  def set_closed_mm(closed_mm, gripper_socket):
      gripper_closed_mm[to_num(gripper_socket) - 1] = closed_mm
  end

  def set_open_mm(open_mm, gripper_socket):
      gripper_open_mm[to_num(gripper_socket) - 1] = open_mm
  end

  def gripper_to_mm(value_gripper, gripper_socket):
      closed_norm = get_closed_norm(gripper_socket)
      open_norm = get_open_norm(gripper_socket)
      closed_mm = get_closed_mm(gripper_socket)
      open_mm = get_open_mm(gripper_socket)

      value_norm = (value_gripper / 255) * 100

      slope = (closed_mm - open_mm) / (closed_norm - open_norm)
      value_mm = slope * (value_norm - closed_norm) + closed_mm

      if (value_mm > open_mm):
          value_mm_limited = open_mm
      elif (value_mm < closed_mm):
          value_mm_limited = closed_mm
      else:
          value_mm_limited = value_mm
      end

      return value_mm_limited
  end

  def mm_to_gripper(value_mm, gripper_socket):
      closed_norm = get_closed_norm(gripper_socket)
      open_norm = get_open_norm(gripper_socket)
      closed_mm = get_closed_mm(gripper_socket)
      open_mm = get_open_mm(gripper_socket)

      slope = (closed_norm - open_norm) / (closed_mm - open_mm)
      value_norm = (value_mm - closed_mm) * slope + closed_norm

      value_gripper = value_norm * 255 / 100

      if (value_gripper > 255):
          value_gripper_limited = 255
      elif (value_gripper < 0):
          value_gripper_limited = 0
      else:
          value_gripper_limited = round_value(value_gripper)
      end

      return value_gripper_limited
  end

  def round_value(value):
      value_mod = value % 1

      if(value_mod < 0.5):
          return floor(value)
      else:
          return ceil(value)
      end
  end

  def round_value_2_dec(value):
      value_x_100 = value * 100
      value_x_100_rounded = round_value(value_x_100)
      return value_x_100_rounded / 100
  end

  def clear_socket_buffer(gripper_socket="1", read_timeout = 0.1):
      rq_comm_clear_socket_buffer_enabled[rq_socket_to_index(gripper_socket)] = True
  end

  def rq_gripper_id_to_ascii(gripper_id):
      if(gripper_id == "1"):
          return 57
      elif(gripper_id == "2"):
          return 50
      elif(gripper_id == "3"):
          return 51
      elif(gripper_id == "4"):
          return 52
      end
  end

      def scale(value, rawRange, scaledRange):
          def computeSlope(inputRange, outputRange):
              outputRangeDelta = outputRange[1] - outputRange[0]
              inputRangeDelta = inputRange[1] - inputRange[0]

              if (inputRangeDelta == 0):
                  return 0
              else:
                  return outputRangeDelta / inputRangeDelta
              end
          end

          def computeIntercept(slope, inputRange, outputRange):
              return outputRange[0] - (slope * inputRange[0])
          end

          def clipScaledValue(outputScaledValue, outputRange):
              if (outputRange[0] < outputRange[1]):
                  return clipWhenLowerLimitIsLessThanHigher(outputScaledValue, outputRange)
              else:
                  return clipWhenLowerLimitIsGreaterThanHigherLimit(outputScaledValue, outputRange)
              end
          end

          def clipWhenLowerLimitIsGreaterThanHigherLimit(outputScaledValue, outputRange):
              if (outputScaledValue < outputRange[1]):
                  return outputRange[1]
              elif (outputScaledValue > outputRange[0]):
                  return outputRange[0]
              else:
                  return outputScaledValue
              end
          end

          def clipWhenLowerLimitIsLessThanHigher(outputScaledValue, outputRange):
              if (outputScaledValue < outputRange[0]):
                  return outputRange[0]
              elif (outputScaledValue > outputRange[1]):
                  return outputRange[1]
              else:
                  return outputScaledValue
              end
          end

          slope = computeSlope(rawRange, scaledRange)
          intercept = computeIntercept(slope, rawRange, scaledRange)
          scaledValue = slope * value + intercept
          return clipScaledValue(scaledValue, scaledRange)
      end

      def limit(value, range):
          return scale(value, range, range)
      end


  rq_init_comm_if_connected(9, "1")
  rq_init_comm_if_connected(2, "2")
  rq_init_comm_if_connected(3, "3")
  rq_init_comm_if_connected(4, "4")
  rq_print_connected_grippers()
  rq_gripper_communication_thread = run rq_gripper_communication()
  set_closed_norm(97.6470588235294, "1")
  set_open_norm(1.1764705882352942, "1")
  set_closed_mm(0.0, "1")
  set_open_mm(53.0, "1")
  set_closed_norm(100.0, "2")
  set_open_norm(0.0, "2")
  set_closed_mm(0.0, "2")
  set_open_mm(50.0, "2")
  set_closed_norm(100.0, "3")
  set_open_norm(0.0, "3")
  set_closed_mm(0.0, "3")
  set_open_mm(50.0, "3")
  set_closed_norm(100.0, "4")
  set_open_norm(0.0, "4")
  set_closed_mm(0.0, "4")
  set_open_mm(50.0, "4")
  rq_current_limit_enabled = False
  while(not rq_gripper_communication_thread_started):
      sleep(0.008)
  end
  # end: URCap Installation Node
  global AMR_Position=struct(position_identifier=0, x1=0, x2=0, y1=0, y2=0, theta1=0, theta2=0)
  global CAM_Pose=p[0,0,0,0,0,0]
  global CAM_Relation=""
  global CMD_Abort=  False
  global CMD_Clear=  False
  global CMD_Reset=  False
  global CMD_Start=  False
  global CMD_Suspend=  False
  global CMD_Unhold=  False
  global CMD_Unsuspend=  False
  global CNT_Rack_Output=0
  global FNC_Freedrive=  False
  global PRC_TubCounter=0
  global STP=0
  global easyPickCount_4=0
  global easyPickCount_7=0
  global easyPickNoObj_4=0
  global easyPickNoObj_7=0
  global easyPickParts_4=0
  global easyPickParts_7=0
  global TMR_Barcode=0
  global Container_mid_1_p=p[-.379239199143, -.127191311915, .299999999998, .000000000046, -.000000000021, -1.247199999994]
  global Container_mid_1_q=[-2.477408934449926, -1.2969853503591224, -1.875639182904262, -1.539621866126728, 1.5731943360401213, -2.8009955944022717]
  global trigger_otw_p=p[-.364831738276, -.163967193938, .343299997821, .000000000046, -.000000000020, -1.148401333327]
  global trigger_otw_q=[-2.378283213085033, -1.2994862387706814, -1.7634300687554951, -1.6493302004167063, 1.573123683454141, -2.8011223671816943]
  global Waypoint_54_p=p[.008800512419, -.547926542621, .402696567415, -.589884378425, -.007228654778, -.061268144704]
  global Waypoint_54_q=[-1.2044575850116175, -1.3416667741588135, -1.8272563219070435, -0.9884541195682068, 1.3621035814285278, -2.7712565104113978]
  global Waypoint_77_p=p[-.178371829612, -.433927395311, .368082383916, -.086593488055, .704679941724, -.007869906074]
  global Waypoint_77_q=[-1.265390698109762, -1.3355963987163086, -1.7944865226745605, -1.7402602634825648, 0.8780410885810852, -2.7713127771960657]
  global Waypoint_83_p=p[.008800512419, -.547926542621, .402696567415, -.589884378425, -.007228654778, -.061268144704]
  global Waypoint_83_q=[-1.2044575850116175, -1.3416667741588135, -1.8272563219070435, -0.9884541195682068, 1.3621035814285278, -2.7712565104113978]
  global Waypoint_84_p=p[-.178371829612, -.433927395311, .368082383916, -.086593488055, .704679941724, -.007869906074]
  global Waypoint_84_q=[-1.265390698109762, -1.3355963987163086, -1.7944865226745605, -1.7402602634825648, 0.8780410885810852, -2.7713127771960657]
  global Vial_above_1_p=p[.017105793010, -.652093028359, .184920586844, .000000000272, .000000000270, 1.564063451276]
  global Vial_above_1_q=[-1.3375440709712851, -1.9618096977868804, -1.4665759083780685, -1.2837941559171444, 1.5732503672317195, -4.47276330421513]
  global Vial_pick_poi_1_p=p[.017105792852, -.648922724010, .093307568731, .000000000271, .000000000270, 1.564063451276]
  global Vial_pick_poi_1_q=[-1.3366329456391917, -2.0375277831965413, -1.6071432798879028, -1.0675084332049813, 1.57309887265915, -4.471135348858068]
  global Waypoint_86_p=p[.019227646885, -.648669633640, .184920586950, .000000000000, .000000000000, .024063451426]
  global Waypoint_86_q=[-1.3331129109407733, -1.9540750545686123, -1.4775914902901128, -1.280581784992414, 1.5733500744865856, -2.928303704452631]
  global Waypoint_87_p=p[-.032361834699, -.348336136197, .391475576335, -.000008499254, .000014589902, -.004651426820]
  global Waypoint_87_q=[-1.2709335019096129, -1.1914598663441005, -1.708995335060501, -1.8117888533498316, 1.5729683532263925, -2.8379347397710237]
  global Vial_3FG_plac_1_p=p[-.031858676359, -.349402499566, .145301120695, .000000000000, .000000000000, .000000000000]
  global Vial_3FG_plac_1_q=[-1.2723975525801707, -1.252376585823825, -2.3128114007049496, -1.1470592278900167, 1.5730548099411423, -2.8414815174610535]
  global Waypoint_88_p=p[-.032361834699, -.348336136197, .391475576335, -.000008499254, .000014589902, -.004651426820]
  global Waypoint_88_q=[-1.2709335019096129, -1.1914598663441005, -1.708995335060501, -1.8117888533498316, 1.5729683532263925, -2.8379347397710237]
  global cap_dump_1_p=p[-.139168676487, -.420163541420, .146096395183, .000000000000, .000000000000, .000000000000]
  global cap_dump_1_q=[-1.584588644510994, -1.5093464179777323, -2.1118449369620347, -1.091059703602438, 1.5728943834877336, -3.154014906686923]
  global Waypoint_89_p=p[-.032361834699, -.348336136197, .391475576335, -.000008499254, .000014589902, -.004651426820]
  global Waypoint_89_q=[-1.2709335019096129, -1.1914598663441005, -1.708995335060501, -1.8117888533498316, 1.5729683532263925, -2.8379347397710237]
  global Vial_3FG_plac_2_p=p[-.031858676359, -.349402499566, .145301120695, .000000000000, .000000000000, .000000000000]
  global Vial_3FG_plac_2_q=[-1.2723975525801707, -1.252376585823825, -2.3128114007049496, -1.1470592278900167, 1.5730548099411423, -2.8414815174610535]
  global Waypoint_90_p=p[-.032361834699, -.348336136197, .391475576335, -.000008499254, .000014589902, -.004651426820]
  global Waypoint_90_q=[-1.2709335019096129, -1.1914598663441005, -1.708995335060501, -1.8117888533498316, 1.5729683532263925, -2.8379347397710237]
  global cap_dump_2_p=p[-.139168676487, -.420163541420, .146096395183, .000000000000, .000000000000, .000000000000]
  global cap_dump_2_q=[-1.584588644510994, -1.5093464179777323, -2.1118449369620347, -1.091059703602438, 1.5728943834877336, -3.154014906686923]
  global Waypoint_91_p=p[-.032361834699, -.348336136197, .391475576335, -.000008499254, .000014589902, -.004651426820]
  global Waypoint_91_q=[-1.2709335019096129, -1.1914598663441005, -1.708995335060501, -1.8117888533498316, 1.5729683532263925, -2.8379347397710237]
  global Vial_liq_abov_1_p=p[-.025303660977, -.338758622354, .426628485936, -1.315858642253, .800043520260, -.928295855026]
  global Vial_liq_abov_1_q=[-0.3789628187762659, -1.5149522957256814, -2.263045310974121, 0.7870649534412841, -0.750984017048971, -3.2237566153155726]
  global Vial_liq_pick_3_p=p[-.002660428945, -.335984893034, .159389832934, -1.150456778400, .673175527684, -1.010612657503]
  global Vial_liq_pick_3_q=[-0.3660772482501429, -1.4503649038127442, -2.4056053161621094, -1.994692941705221, 0.8039668202400208, -0.2508929411517542]
  global Vial_liq_pick_4_p=p[-.041402486291, -.356791603314, .125395323246, -1.143483969075, .651070210027, -.878721885453]
  global Vial_liq_pick_4_q=[-0.4426233705502476, -1.437252121513727, -2.551930962114307, -1.776528229806984, 0.6562026234073748, -0.43018811960029524]
  global Vial_liq_abov_2_p=p[-.025303660977, -.338758622354, .426628485936, -1.315858642253, .800043520260, -.928295855026]
  global Vial_liq_abov_2_q=[-0.3789628187762659, -1.5149522957256814, -2.263045310974121, 0.7870649534412841, -0.750984017048971, -3.2237566153155726]
  global Liquid_midway_1_p=p[.057575295009, -.583081747994, .306414980749, -1.351675548728, .120935756539, -.096908606303]
  global Liquid_midway_1_q=[-0.895174805318014, -1.7035466633238734, -2.380953073501587, 0.631549521083496, 0.7706599235534668, -2.9455552736865442]
  global shake_3_p=p[.057574880217, -.583085370269, .306422893466, -1.360996190983, -.155555042453, -.438136255921]
  global shake_3_q=[-0.8951800505267542, -1.7035466633238734, -2.380937099456787, 0.6315542894550782, 0.7706599235534669, -2.5394540616517496]
  global shake_4_p=p[.057581636113, -.583090570002, .306439684073, -1.308767904323, .368530312677, .214926493520]
  global shake_4_q=[-0.8951714674579065, -1.7035395107665003, -2.380906343460083, 0.6315504747578125, 0.7706480026245118, -3.3161255787892268]
  global drop_above_3_p=p[.268235025993, -.467784390499, .226219872376, -1.027832627524, -.430841408251, 1.004603115937]
  global drop_above_3_q=[-0.935645882283346, -1.6663371525206507, -2.4252893924713135, 0.41966931402172847, 1.8470635414123535, -3.4600217978106897]
  global drop_above_4_p=p[.219042229014, -.470775657081, .133754190740, -.313004595901, -.344395319364, 1.500564994056]
  global drop_above_4_q=[-1.0601594887284795, -1.70046459045642, -2.0799996233759863, -0.7243227230676759, 1.9429634314685202, -4.115129153870795]
  global liq_tran_3_p=p[.213067510942, -.469567035397, .100231043184, .251862243732, .217902579404, 1.592812335393]
  global liq_tran_3_q=[-0.7789645168037476, -1.822364827406652, -1.8643518410805573, -1.252158963840138, 1.3768134449520435, -3.9328333233290254]
  global drop_above_5_p=p[.219042229014, -.470775657081, .133754190740, -.313004595901, -.344395319364, 1.500564994056]
  global drop_above_5_q=[-1.0601594887284795, -1.70046459045642, -2.0799996233759863, -0.7243227230676759, 1.9429634314685202, -4.115129153870795]
  global Waypoint_92_p=p[.187119460405, -.493959476151, .133754190608, -.313004596540, -.344395317757, 1.500564993991]
  global Waypoint_92_q=[-1.1418328121400876, -1.7310553375189475, -2.033634768766424, -0.772026910513711, 1.958578934631971, -4.201588449364511]
  global liq_tran_4_p=p[.195957706507, -.493022614126, .100231042689, .160718757180, .109807038912, 1.525321508623]
  global liq_tran_4_q=[-0.881740380645474, -1.8244526267589851, -1.865100964490387, -1.1608866323693583, 1.4631433601076713, -3.973915130363038]
  global drop_above_6_p=p[.219042229014, -.470775657081, .133754190740, -.313004595901, -.344395319364, 1.500564994056]
  global drop_above_6_q=[-1.0601594887284795, -1.70046459045642, -2.0799996233759863, -0.7243227230676759, 1.9429634314685202, -4.115129153870795]
  global drop_above_7_p=p[.268235025993, -.467784390499, .226219872376, -1.027832627524, -.430841408251, 1.004603115937]
  global drop_above_7_q=[-0.935645882283346, -1.6663371525206507, -2.4252893924713135, 0.41966931402172847, 1.8470635414123535, -3.4600217978106897]
  global Liquid_midway_2_p=p[.057575295009, -.583081747994, .306414980749, -1.351675548728, .120935756539, -.096908606303]
  global Liquid_midway_2_q=[-0.895174805318014, -1.7035466633238734, -2.380953073501587, 0.631549521083496, 0.7706599235534668, -2.9455552736865442]
  global Vial_drop_abo_1_p=p[.000324902251, -.648569523142, .221894115667, -.873462921366, 1.165852672573, -1.482720593185]
  global Vial_drop_abo_1_q=[-1.0576906334721352, -2.393016994184633, -0.9236232851859159, -2.5729213042279273, 0.7903331288549689, -0.33286325848155585]
  global Vial_liq_drop_1_p=p[.001020867953, -.647659915585, .092915870838, -.834762611599, 1.081942994823, -1.540647900176]
  global Vial_liq_drop_1_q=[-1.0631954168193474, -2.4447642951220825, -1.128811017825127, -2.1983115491972294, 0.8130148661460634, -0.38984988696911316]
  global Vial_drop_abo_2_p=p[.000324902251, -.648569523142, .221894115667, -.873462921366, 1.165852672573, -1.482720593185]
  global Vial_drop_abo_2_q=[-1.0576906334721352, -2.393016994184633, -0.9236232851859159, -2.5729213042279273, 0.7903331288549689, -0.33286325848155585]
  global Spatula_otw_p=p[-.038472058237, -.263141484147, .425351216717, -.000441582511, -.000128175490, 3.034387645854]
  global Spatula_otw_q=[-1.1888947506684495, -1.0083288774886814, -1.7052227056065874, -1.9984805067363443, 1.5730180972985317, 0.48793409320312264]
  global pick_spat_L_abv_p=p[.239059466375, -.067212518441, .280720723617, .000017217488, -.000484427718, 3.106837214660]
  global pick_spat_L_abv_q=[0.292765616142962, -0.8565557553273315, -2.140199892763044, -1.715349495646084, 1.573623142106424, 1.8984976776985687]
  global spat_L_pick_p=p[.242468789885, -.067301915011, .193171208067, .000017217488, -.000484427718, 3.106837214657]
  global spat_L_pick_q=[0.2867414378807389, -0.8600077002089179, -2.3629148016312627, -1.4891831672860159, 1.5737695566221115, 1.8933890858591198]
  global spat_L_lift_p=p[.245402002494, -.067432373551, .289049296496, .000017217490, -.000484427724, 3.106837214657]
  global spat_L_lift_q=[0.2834351187564135, -0.8798320076811592, -2.1119436738532986, -1.7203314352121302, 1.573588313403067, 1.8891054681654005]
  global spat_L_side_p=p[.247133573905, -.017633681797, .289062935631, .000017217490, -.000484427724, 3.106837214657]
  global spat_L_side_q=[0.49719173575848863, -0.8582398211168538, -2.1182130454788215, -1.735610316654931, 1.5735817737572706, 2.1028402698705397]
  global spat_L_up_p=p[.247135508891, -.017665229117, .420978991173, .000017217478, -.000484427734, 3.106837214657]
  global spat_L_up_q=[0.4989125281866238, -0.9581229935107345, -1.7344014311356126, -2.0195384609726084, 1.5729657310403162, 2.10331546461867]
  global spat_M_up_p=p[.244553462372, -.113574254431, .420343304672, .000026293938, -.000477463024, 3.067686801419]
  global spat_M_up_q=[0.08431285927297782, -1.0128123619317435, -1.7175182391153623, -1.9818233355759816, 1.5730135231275326, 1.727892677465693]
  global spat_M_pick_p=p[.244642228055, -.114374053673, .192299012591, .000045577878, -.000000729326, 3.128037167562]
  global spat_M_pick_q=[0.07853961211226647, -0.930778014039741, -2.3425698873551504, -1.4388489853835722, 1.5733856270317392, 1.6640658846527625]
  global spat_S_Up_7_p=p[.243228810603, -.161948321982, .423281604617, .000026293955, -.000477463064, 3.067686800854]
  global spat_S_Up_7_q=[-0.11182322368059516, -1.0716267311491734, -1.6854498186860427, -1.955120134033855, 1.5730106579635699, 1.5317349120701778]
  global spat_S_Pick_4_p=p[.245377020686, -.158668022535, .192285730279, .000026293986, -.000477463054, 3.127999999999]
  global spat_S_Pick_4_q=[-0.10086534461938079, -1.0111878731926387, -2.3119775963829685, -1.3890307323937048, 1.5735923824164428, 1.4847497788366055]
  global spat_S_Up_8_p=p[.252087445596, -.159242094834, .423281604617, .000026293954, -.000477463070, 3.067686800855]
  global spat_S_Up_8_q=[-0.09804692328730358, -1.0862987822056382, -1.6788706463996483, -1.9470242450550348, 1.5730147401359813, 1.5455107082823842]
  global spat_flatM_up_p=p[.241028517126, -.208127630016, .404671074680, .000026293951, -.000477463078, 3.067686800891]
  global spat_flatM_up_q=[-0.27878462628263456, -1.1217510366315881, -1.7121530048618725, -1.8783279876432832, 1.5731053960668042, 1.3649536117980254]
  global spat_flatM_pick_p=p[.241028983327, -.208057297586, .192270533170, .000026293950, -.000477463079, 3.067686800885]
  global spat_flatM_pick_q=[-0.2805687960562633, -1.1003763929487214, -2.271431297337675, -1.3404236887924883, 1.5734924238720627, 1.3653813047742556]
  global spat_flatS_up_p=p[.237651953780, -.253943828614, .403961222825, .000026293950, -.000477463092, 3.067686800841]
  global spat_flatS_up_q=[-0.42363550926974103, -1.1939944599502539, -1.6745915127240307, -1.843675057902054, 1.5731001874678698, 1.220082820532415]
  global spat_flatS_pick_p=p[.241325662334, -.251726327528, .192256842740, .000026293947, -.000477463087, 3.067686800841]
  global spat_flatS_pick_q=[-0.4144907797170738, -1.1967447109013012, -2.21926362252748, -1.2962499335425761, 1.5733885098427622, 1.2314402238866728]
  global spat_S_pick_p=p[.241585614619, -.158882677087, .191636172448, .000019478956, -.000483249177, 3.097147973434]
  global spat_S_pick_q=[-0.10320942227973173, -1.0007485193115802, -2.317947069452162, -1.3934956127505886, 1.5736112980229278, 1.5132597021160705]
  global spat_S_up_p=p[.248189103503, -.159371150053, .417088864416, .000026293966, -.000477463070, 3.067686800840]
  global spat_S_up_q=[-0.10007737460061872, -1.0730270029702904, -1.7018049146034766, -1.9373622285571734, 1.573045444550866, 1.5435422173047084]
  global Waypoint_7_p=p[-.472820924474, .292439826233, .207418370237, -.137787250486, 2.177332259632, -2.152029714756]
  global Waypoint_7_q=[-2.911134078210732, -1.90240864358569, -1.968768330510411, -2.500365101593811, 0.11427687110891149, 0.0958980389250167]
  global Waypoint_8_p=p[-.357612884176, -.251084817998, .212379799667, -.858181193174, 1.714832512191, -1.687547565568]
  global Waypoint_8_q=[-1.620834863369681, -1.8936194567376496, -1.9821394403832038, -2.4599791457905273, 0.6296693672615152, 0.07625365420707819]
  global Decapp_above_3_p=p[-.013480295948, -.359153355979, .266194408367, -.879653555922, 1.646336924805, -1.709111068605]
  global Decapp_above_3_q=[-0.9632157249872035, -2.0163405763031657, -1.5968194594157152, -2.6579215719847085, 1.251243398585566, 0.047906446502667066]
  global Decapp_place_3_p=p[-.013480295890, -.359153356055, .160907502384, -.879653554902, 1.646336919740, -1.709111066456]
  global Decapp_place_3_q=[-0.9633402410919709, -2.1541179572356635, -1.6937729380888573, -2.4232786481058053, 1.2517342187662468, 0.04818402956922263]
  global Decapp_above_4_p=p[-.013480295948, -.359153355979, .266194408367, -.879653555922, 1.646336924805, -1.709111068605]
  global Decapp_above_4_q=[-0.9632157249872035, -2.0163405763031657, -1.5968194594157152, -2.6579215719847085, 1.251243398585566, 0.047906446502667066]
  global Waypoint_78_p=p[-.051450028091, -.519555688329, .365718563414, -1.287302938145, 1.077637394477, -1.218524965834]
  global Waypoint_78_q=[-0.9214276262416012, -1.8899696965062578, -1.4939326452510562, -2.840015661555725, 0.5585157189668353, 0.033997638875617575]
  global Waypoint_10_p=p[-.466751210260, .252836712095, .259921246286, 1.042686976164, .439333316918, -1.691967798809]
  global Waypoint_10_q=[-3.022216346250036, -1.8383597675135919, -1.566977059184386, -2.046864464116096, 0.8487467526238, -2.4392912369481916]
  global Waypoint_9_p=p[-.538777454962, .370695704977, .175030018143, -.317104215445, 2.082346543003, -2.037631421082]
  global Waypoint_9_q=[-3.1158871966457857, -1.998548595120492, -1.941797010061462, -2.2703530575838844, -0.27573365931009164, -0.06926782177267654]
  global Powder_wayp1_p=p[-.472820924474, .292439826233, .207418370237, -.137787250486, 2.177332259632, -2.152029714756]
  global Powder_wayp1_q=[-2.911134078210732, -1.90240864358569, -1.968768330510411, -2.500365101593811, 0.11427687110891149, 0.0958980389250167]
  global Waypoint_2_p=p[-.357612884176, -.251084817998, .212379799667, -.858181193174, 1.714832512191, -1.687547565568]
  global Waypoint_2_q=[-1.620834863369681, -1.8936194567376496, -1.9821394403832038, -2.4599791457905273, 0.6296693672615152, 0.07625365420707819]
  global Postions_otw_p=p[-.010896578244, -.533368729951, .288851175116, -1.233738470894, 1.195331112012, -1.207314088469]
  global Postions_otw_q=[-0.898791023514228, -2.078490033037677, -1.4499891355755317, -2.7624416226992476, 0.6570218891920963, 0.02136606178275929]
  global cont_A_otw_p=p[.070238108556, -.655257851554, .184611566008, -1.090601381517, 1.404822685081, -1.413645380264]
  global cont_A_otw_q=[-0.990969136335913, -2.7123780097559784, -0.5772671651193146, -3.0005537851220403, 0.84719335943793, 0.020652463706785973]
  global cont_B_otw_p=p[.255895686750, -.501120003087, .157855243207, -1.209177187561, 1.209243088037, -1.209202949417]
  global cont_B_otw_q=[-0.5819602570351563, -2.5181180937953833, -1.0264696604583161, -2.7360726814058687, 0.9880932038785559, -0.004134033524621827]
  global cont_B_safe_p=p[.242897168204, -.501733713795, .237745474779, -1.209212324107, 1.209144328638, -1.209309913894]
  global cont_B_safe_q=[-0.5929699566143585, -2.4210115429142114, -0.9949203644592259, -2.8646436479104267, 0.976678899749076, -0.004020526358775811]
  global cont_C_otw_p=p[.319495487998, -.362719410364, .163846736977, -1.233784872294, 1.195277203291, -1.207325031551]
  global cont_C_otw_q=[-0.3611889651645974, -2.404603865546651, -1.2341573845076566, -2.650535279811077, 1.1944844573128257, 0.01638086594640864]
  global Waypoint_1_p=p[-.352029261722, -.424157832422, .472326578019, -.000004407962, .000020663369, -1.529709227737]
  global Waypoint_1_q=[-2.017015745614491, -1.7423968528991196, -1.0053357238485425, -1.9644715035904907, 1.5727249689896, -2.060727852912713]
  global Waypoint_5_p=p[.219993437017, -.447144142811, .462350040687, .000006087494, .000031090075, .000022232405]
  global Waypoint_5_q=[-0.8406239476037944, -1.5982534362206806, -1.1934200873248484, -1.9205794898315975, 1.5727336676986443, -2.4135960466995314]
  global place_2_home_p=p[-.352029261717, -.424157832411, .329197314759, -.000004407962, .000020663369, -1.529709227737]
  global place_2_home_q=[-2.017880982348384, -1.6708952803108668, -1.462293789471877, -1.5790150659586653, 1.5732060241635952, -2.059940179665328]
  global Waypoint_12_p=p[-.812560029877, -.415067232840, .258518340146, -1.257569567036, 1.159670338548, -1.145019586130]
  global Waypoint_12_q=[-2.3224548809497123, -2.3211405271930765, -1.1304722687551445, -2.8155296475017018, -0.8321758827962036, -0.007205995478960503]
  global Waypoint_18_p=p[-.813643087636, -.416224939441, .099970000000, -1.257570310935, 1.159676546330, -1.145010619029]
  global Waypoint_18_q=[-2.322494764677227, -2.501268559301314, -1.239250885783676, -2.5265468980680197, -0.831327849164623, -0.00732105677136996]
  global Waypoint_19_p=p[-.812560029269, -.415067232191, .079455005744, -1.257569567033, 1.159670338546, -1.145019586137]
  global Waypoint_19_q=[-2.3224951834453367, -2.5274729453886575, -1.2489176533831348, -2.4906644180980346, -0.8312252662037514, -0.007338111970053518]
  global Scan_db_p=p[-.000000000035, -.399999999894, .423061661675, .000000000000, .000000000000, .000000000000]
  global Scan_db_q=[-1.2292165564781996, -1.3327911122625213, -1.5324793532106682, -1.846975993436244, 1.5728640135188283, -2.801307704234451]
  global TMR_Barcode_is_counting=False
  thread Timer_Thread():
    while (True):
      if (TMR_Barcode_is_counting):
        TMR_Barcode = TMR_Barcode + get_steptime()
      end
      sync()
    end
  end
  run Timer_Thread()
  def Sub_Vision_V18():
    $ 900 "Sub_Vision_V18" "noBreak"
    $ 901 "PreSettings"
    $ 902 "CAM_LM_Detected≔ False "
    global CAM_LM_Detected=  False
    $ 903 "CAM_Captures≔0"
    global CAM_Captures=0
    $ 904 "CAM_Pose≔p[0,0,0,0,0,0]"
    global CAM_Pose=p[0,0,0,0,0,0]
    $ 905 "CAM_LM_Refinmnt≔ False "
    global CAM_LM_Refinmnt=  False
    $ 906 "CAM_LM_Refined≔ False "
    global CAM_LM_Refined=  False
    $ 907 "CAM_LM_Deviatn≔p[0,0,0,0,0,0]"
    global CAM_LM_Deviatn=p[0,0,0,0,0,0]
    $ 908 "CAM_LM_ID≔0"
    global CAM_LM_ID=0
    $ 909 "CAM_Done≔ False "
    global CAM_Done=  False
    $ 910 "CAM_CNT_Obj≔0"
    global CAM_CNT_Obj=0
    $ 911 "CAM_Result = []"
    CAM_Result = []
    $ 912 "OBJ_Detected≔ False "
    global OBJ_Detected=  False
    $ 913 "FRM_Reference≔p[0,0,0,0,0,0]"
    global FRM_Reference=p[0,0,0,0,0,0]
    $ 914 "'=========='"
    # '=========='
    $ 915 "Switch Action"
    switch_1 = Action
    $ 916 "Case 13"
    if (13 == switch_1):
    elif (15 == switch_1):
      $ 1034 "Case 15"
    elif (131 == switch_1):
      $ 1080 "Case 131"
      $ 1081 "Read (SensoPart)"
      $ 1082 "Action_Info≔'search for landmark'"
      global Action_Info="search for landmark"
      $ 1083 "CAM_LM≔CAM_LMs[4]"
      global CAM_LM=CAM_LMs[4]
      $ 1084 "CAM_Relation≔CAM_LM.capture_relation"
      global CAM_Relation=CAM_LM.capture_relation
      $ 1085 "go to capture pose"
      $ 1088 "If ITM_ID≟1 and JIG≟7"
      if (ITM_ID == 1  and  JIG == 7):
        $ 1089 "PSE_T≔uLM_Cap_SSRack"
        global PSE_T=uLM_Cap_SSRack
      else:
        $ 1090 "ElseIf ITM_ID≟5 and JIG≟7"
        if (ITM_ID == 5  and  JIG == 7):
          $ 1091 "PSE_T≔FRM_Cap_SSRack"
          global PSE_T=FRM_Cap_SSRack
        else:
          $ 1094 "ElseIf ITM_ID≟1 and JIG≟15"
          if (ITM_ID == 1 and JIG == 15):
            $ 1095 "MoveJ"
            $ 1096 "Container_mid_1" "breakAfter"
            movej(get_inverse_kin(Container_mid_1_p, qnear=Container_mid_1_q), a=1.3962634015954636, v=1.0471975511965976, r=0.05)
            $ 1098 "PSE_T≔FRM_Container_const"
            global PSE_T=p[-0.5003348223692186,0.35061804815168285,0.41579001388808423,-5.092943187272062E-5,1.0145185065363121E-4,-2.764319258713288]
          else:
            $ 1099 "ElseIf ITM_ID≟1 and JIG≟21"
            if (ITM_ID == 1 and JIG == 21):
              $ 1100 "Set"
              set_tcp(p[0.0,0.0,0.15052000000000001,3.1415,0.0,0.0])
              $ 1101 "PSE_T≔FRM_PoTS_const"
              global PSE_T=p[-0.5403054403210852,-0.10910773999775857,0.4828,3.058497512721046E-6,2.3454853329357316E-5,-2.208510541952706]
            else:
              $ 1102 "ElseIf ITM_ID≟1 and JIG≟17"
              if (ITM_ID == 1 and JIG == 17):
                $ 1103 "MoveJ"
                $ 1104 "zero_scale()"
                zero_scale()
                $ 1105 "trigger_otw" "breakAfter"
                movej(get_inverse_kin(trigger_otw_p, qnear=trigger_otw_q), a=1.3962634015954636, v=1.0471975511965976, r=0.05)
                $ 1109 "PSE_T≔FRM_weigh_scale_const"
                global PSE_T=p[-0.3804866881697204,0.025744252835212,0.4723487455232425,-1.0445769542396123E-4,-1.924788411074358E-5,-2.1691978730572363]
              end
            end
          end
        end
      end
      $ 1110 "do_transition(PSE_T, keep_rxry=False)"
      do_transition(PSE_T, keep_rxry=False)
      $ 1111 "Set"
      set_tcp(p[0.0,0.0,0.161,3.1415,0.0,0.0])
      $ 1112 "MoveJ"
      $ 1113 "PSE_T" "breakAfter"
      movej(PSE_T, a=1.3962634015954636, v=1.7453292519943295)
      $ 1114 "CAM_Pose≔get_actual_tcp_pose()"
      global CAM_Pose= get_actual_tcp_pose ()
      $ 1115 "Loop  not CAM_Done and  not ERROR.FLAG and  not CMD_Stop"
      while (  not  CAM_Done  and    not  ERROR.FLAG  and    not  CMD_Stop):
        $ 1116 "adjust capture pose"
        $ 1117 "If CAM_LM_Detected and CAM_LM_Refinmnt"
        if (CAM_LM_Detected  and  CAM_LM_Refinmnt):
          $ 1118 "PSE_T≔p[0,0,0.300,0,0,0]"
          global PSE_T=p[0,0,0.300,0,0,0]
          $ 1119 "CAM_Pose≔PSE_T"
          global CAM_Pose=PSE_T
          $ 1120 "If  not is_reachable(FRM_Reference,[PSE_T])"
          if (  not  is_reachable(FRM_Reference,[PSE_T])):
            $ 1121 "Error"
            $ 1122 "set_error(ERROR_POSE_NOT_REACHABLE)"
            set_error(ERROR_POSE_NOT_REACHABLE)
          end
          $ 1123 "If  not ERROR.FLAG"
          if (  not  ERROR.FLAG):
            $ 1124 "MoveJ"
            $ 1125 "PSE_T" "breakAfter"
            set_tcp(p[0.0,0.0,0.161,0.0,0.0,0.0])
            movej(pose_trans(FRM_Reference, PSE_T), a=0.8726646259971648, v=1.3962634015954636)
            $ 1126 "CAM_LM_Refined≔ True "
            global CAM_LM_Refined=  True
          end
        else:
          $ 1127 "ElseIf  not CAM_LM_Detected and CAM_Captures>0"
          if (  not  CAM_LM_Detected  and  CAM_Captures>0):
            $ 1128 "MoveL"
            $ 1129 "If FRM_Reference≟p[0,0,0,0,0,0]"
            if (FRM_Reference == p[0,0,0,0,0,0]):
              $ 1130 "PSE_T≔get_random_pose(pose_ref=CAM_Pose, mode='cubic', range_max=[0.150,0.150,0.015])"
              global PSE_T=get_random_pose(pose_ref=CAM_Pose, mode="cubic", range_max=[0.150,0.150,0.015])
            else:
              $ 1135 "Else" "noBreak"
              $ 1136 "PSE_T≔get_random_pose(pose_ref=CAM_Pose, mode='rotation', range_max=[10,10,0])"
              global PSE_T=get_random_pose(pose_ref=CAM_Pose, mode="rotation", range_max=[10,10,0])
              $ 1137 "CAM_LM_Refined≔ True "
              global CAM_LM_Refined=  True
            end
            $ 1138 "If get_inverse_kin_has_solution(pose_trans(FRM_Reference, PSE_T))"
            if (get_inverse_kin_has_solution( pose_trans (FRM_Reference, PSE_T))):
              $ 1139 "Comment"
              # Comment
              $ 1140 "PSE_T" "breakAfter"
              set_tcp(p[0.0,0.0,0.161,3.1415,0.0,0.0])
              movel(pose_trans(FRM_Reference, PSE_T), a=0.03, v=0.05)
            else:
              $ 1141 "Else" "noBreak"
              $ 1142 "'If random pose is out of reach, set the initial cam pose'"
              # 'If random pose is out of reach, set the initial cam pose'
              $ 1143 "PSE_T≔CAM_Pose"
              global PSE_T=CAM_Pose
            end
          end
        end
        $ 1144 "Wait: 2.0"
        sleep(2.0)
        $ 1145 "trigger"
        $ 1146 "If ITM_ID≟1 and JIG≟7"
        if (ITM_ID == 1  and  JIG == 7):
          # begin: URCap Program Node
          #   Source: SensoPart VISOR Robotic, 2.0.6, SensoPart Industriesensorik GmbH
          #   Type: VISOR Trigger
          $ 1147 "# 1 VISOR Trigger"
          visor_changeJob(1, "Landmark_INVITE_2", 6000)
          visor_trigger(1, 6000, "arm")
          # end: URCap Program Node
        else:
          $ 1148 "ElseIf ITM_ID≟5 and JIG≟7"
          if (ITM_ID == 5  and  JIG == 7):
            # begin: URCap Program Node
            #   Source: SensoPart VISOR Robotic, 2.0.6, SensoPart Industriesensorik GmbH
            #   Type: VISOR Trigger
            $ 1149 "# 1 VISOR Trigger"
            visor_changeJob(1, "Landmark_INVITE_2", 6000)
            visor_trigger(1, 6000, "arm")
            # end: URCap Program Node
          else:
            $ 1150 "ElseIf ITM_ID≟13 and JIG≟7"
            if (ITM_ID == 13  and  JIG == 7):
              # begin: URCap Program Node
              #   Source: SensoPart VISOR Robotic, 2.0.6, SensoPart Industriesensorik GmbH
              #   Type: VISOR Trigger
              $ 1151 "# 1 VISOR Trigger"
              visor_changeJob(1, "Landmark_INVITE_2", 6000)
              visor_trigger(1, 6000, "arm")
              # end: URCap Program Node
            else:
              $ 1152 "ElseIf ITM_ID≟1 and JIG≟15"
              if (ITM_ID == 1 and JIG == 15):
                # begin: URCap Program Node
                #   Source: SensoPart VISOR Robotic, 2.0.6, SensoPart Industriesensorik GmbH
                #   Type: VISOR Trigger
                $ 1153 "# 1 VISOR Trigger"
                visor_changeJob(1, "Aztec_no_dot_pick", 6000)
                visor_trigger(1, 6000, "arm")
                # end: URCap Program Node
              else:
                $ 1154 "ElseIf ITM_ID≟1 and JIG≟21"
                if (ITM_ID == 1 and JIG == 21):
                  # begin: URCap Program Node
                  #   Source: SensoPart VISOR Robotic, 2.0.6, SensoPart Industriesensorik GmbH
                  #   Type: VISOR Trigger
                  $ 1155 "# 1 VISOR Trigger"
                  visor_changeJob(1, "Fumehood_container", 6000)
                  visor_trigger(1, 6000, "arm")
                  # end: URCap Program Node
                else:
                  $ 1156 "ElseIf ITM_ID≟1 and JIG≟17"
                  if (ITM_ID == 1 and JIG == 17):
                    # begin: URCap Program Node
                    #   Source: SensoPart VISOR Robotic, 2.0.6, SensoPart Industriesensorik GmbH
                    #   Type: VISOR Trigger
                    $ 1157 "# 1 VISOR Trigger"
                    visor_changeJob(1, "Weigh_target", 6000)
                    visor_trigger(1, 6000, "arm")
                    # end: URCap Program Node
                  end
                end
              end
            end
          end
        end
        $ 1161 "TM_3D_Found≔visor_partsFound(1)"
        global TM_3D_Found= visor_partsFound (1)
        $ 1163 "If TM_3D_Found>0"
        if (TM_3D_Found>0):
          $ 1164 "CAM_LM_Detected≔ True "
          global CAM_LM_Detected=  True
          $ 1165 "CAM_Captures≔0"
          global CAM_Captures=0
        else:
          $ 1166 "Else" "noBreak"
          $ 1167 "CAM_LM_Detected≔ False "
          global CAM_LM_Detected=  False
          $ 1168 "CAM_Captures≔CAM_Captures+1"
          global CAM_Captures=CAM_Captures+1
        end
        $ 1173 "result"
        $ 1174 "If CAM_LM_Detected"
        if (CAM_LM_Detected):
          $ 1175 "If (CAM_LM_Refinmnt and CAM_LM_Refined) or  not CAM_LM_Refinmnt"
          if ((CAM_LM_Refinmnt  and  CAM_LM_Refined)  or    not  CAM_LM_Refinmnt):
            $ 1233 "If ITM_ID≟1 and JIG≟7"
            if (ITM_ID == 1  and  JIG == 7):
              $ 1234 "CAM_LM_SSRack≔visor_getPose3d(1, 0)"
              global CAM_LM_SSRack= visor_getPose3d (1, 0)
            else:
              $ 1235 "ElseIf ITM_ID≟5 and JIG≟7"
              if (ITM_ID == 5  and  JIG == 7):
                $ 1236 "CAM_LM_SSRack≔visor_getPose3d(1, 0)"
                global CAM_LM_SSRack= visor_getPose3d (1, 0)
              else:
                $ 1239 "ElseIf ITM_ID≟1 and JIG≟15"
                if (ITM_ID == 1 and JIG == 15):
                  $ 1240 "CAM_LM_cont≔visor_getPose3d(1, 0)"
                  global CAM_LM_cont= visor_getPose3d (1, 0)
                  $ 1241 "Trigger≔get_actual_tcp_pose()"
                  global Trigger= get_actual_tcp_pose ()
                else:
                  $ 1242 "ElseIf ITM_ID≟1 and JIG≟21"
                  if (ITM_ID == 1 and JIG == 21):
                    $ 1243 "CAM_LM_cont≔visor_getPose3d(1, 0)"
                    global CAM_LM_cont= visor_getPose3d (1, 0)
                    $ 1244 "Trigger≔get_actual_tcp_pose()"
                    global Trigger= get_actual_tcp_pose ()
                  else:
                    $ 1245 "ElseIf ITM_ID≟1 and JIG≟17"
                    if (ITM_ID == 1 and JIG == 17):
                      $ 1246 "CAM_LM_cont≔visor_getPose3d(1, 0)"
                      global CAM_LM_cont= visor_getPose3d (1, 0)
                      $ 1247 "Trigger≔get_actual_tcp_pose()"
                      global Trigger= get_actual_tcp_pose ()
                    end
                  end
                end
              end
            end
            $ 1248 "CAM_Done≔ True "
            global CAM_Done=  True
          end
        else:
          $ 1249 "ElseIf  not CAM_LM_Detected and CAM_Captures<CAM_PRM_Retries"
          if (  not  CAM_LM_Detected  and  CAM_Captures<CAM_PRM_Retries):
            $ 1250 "CAM_LM_Refined≔ False "
            global CAM_LM_Refined=  False
          else:
            $ 1251 "ElseIf CAM_Captures≥CAM_PRM_Retries"
            if (CAM_Captures >= CAM_PRM_Retries):
              $ 1252 "CAM_Done≔ True "
              global CAM_Done=  True
              $ 1253 "Error"
              $ 1254 "set_error(ERROR_NO_LANDMARK)"
              set_error(ERROR_NO_LANDMARK)
            end
          end
        end
      end
    elif (151 == switch_1):
      $ 1255 "Case 151"
      $ 1256 "Detect (SensoPart)"
      $ 1257 "go to capture pose"
      $ 1258 "FRM_Reference≔FRM_Cap_SSRack"
      global FRM_Reference=FRM_Cap_SSRack
      $ 1259 "PSE_T≔p[0,0,-0.00,0,0,0]"
      global PSE_T=p[0,0,-0.00,0,0,0]
      $ 1260 "do_transition(pose_trans(FRM_Reference, PSE_T), keep_rxry=False)"
      do_transition( pose_trans (FRM_Reference, PSE_T), keep_rxry=False)
      $ 1261 "JNT_Q≔get_actual_joint_positions()"
      global JNT_Q= get_actual_joint_positions ()
      $ 1262 "JNT_Q≔[JNT_Q[0], JNT_Q[1], JNT_Q[2], JNT_Q[3], JNT_Q[4], 0]"
      global JNT_Q=[JNT_Q[0], JNT_Q[1], JNT_Q[2], JNT_Q[3], JNT_Q[4], 0]
      $ 1263 "Set"
      set_tcp(p[0.0,0.0,0.161,3.1415,0.0,0.0])
      $ 1264 "movej(get_inverse_kin(pose_trans(FRM_Reference, PSE_T), qnear=JNT_Q))"
      movej(get_inverse_kin( pose_trans (FRM_Reference, PSE_T), qnear=JNT_Q))
      $ 1265 "CAM_Pose≔pose_trans(pose_inv(FRM_Reference), get_actual_tcp_pose())"
      global CAM_Pose= pose_trans ( pose_inv (FRM_Reference),  get_actual_tcp_pose ())
      $ 1266 "Loop  not CAM_Done and  not ERROR.FLAG and  not CMD_Stop"
      while (  not  CAM_Done  and    not  ERROR.FLAG  and    not  CMD_Stop):
        $ 1267 "If  not OBJ_Detected and CAM_Captures>0"
        if (  not  OBJ_Detected  and  CAM_Captures>0):
          $ 1268 "MoveL"
          $ 1269 "If FRM_Reference≟p[0,0,0,0,0,0]"
          if (FRM_Reference == p[0,0,0,0,0,0]):
            $ 1271 "PSE_T≔get_random_pose(pose_ref=CAM_Pose, mode='rotation', range_max=[15,15,0])"
            global PSE_T=get_random_pose(pose_ref=CAM_Pose, mode="rotation", range_max=[15,15,0])
          else:
            $ 1272 "Else" "noBreak"
            $ 1273 "PSE_T≔get_random_pose(pose_ref=CAM_Pose, mode='rotation', range_max=[10,10,0])"
            global PSE_T=get_random_pose(pose_ref=CAM_Pose, mode="rotation", range_max=[10,10,0])
          end
          $ 1274 "If get_inverse_kin_has_solution(pose_trans(FRM_Reference, PSE_T))"
          if (get_inverse_kin_has_solution( pose_trans (FRM_Reference, PSE_T))):
            $ 1275 "PSE_T" "breakAfter"
            set_tcp(p[0.0,0.0,0.161,3.1415,0.0,0.0])
            movel(pose_trans(FRM_Reference, PSE_T), a=0.03, v=0.05)
          else:
            $ 1276 "Else" "noBreak"
            $ 1277 "'If random pose is out of reach, set the initial cam pose'"
            # 'If random pose is out of reach, set the initial cam pose'
            $ 1278 "PSE_T≔CAM_Pose"
            global PSE_T=CAM_Pose
            $ 1279 "PSE_T" "breakAfter"
            set_tcp(p[0.0,0.0,0.161,3.1415,0.0,0.0])
            movel(pose_trans(FRM_Reference, PSE_T), a=0.03, v=0.05)
          end
        end
        $ 1280 "Wait: 0.5"
        sleep(0.5)
        $ 1281 "Set"
        set_tcp(p[0.0,0.0,0.161,3.1415,0.0,0.0])
        # begin: URCap Program Node
        #   Source: SensoPart VISOR Robotic, 2.0.6, SensoPart Industriesensorik GmbH
        #   Type: VISOR Trigger
        $ 1282 "# 1 VISOR Trigger"
        visor_changeJob(1, "Object Detection Single", 6000)
        visor_trigger(1, 6000, "arm")
        # end: URCap Program Node
        $ 1283 "If visor_isResponseOk(1)"
        if ( visor_isResponseOk (1)):
          $ 1284 "CAM_CNT_Obj≔visor_partsFound(1)"
          global CAM_CNT_Obj= visor_partsFound (1)
          $ 1285 "CAM_OBJ_Pose≔visor_getPose3d(1, 0)"
          global CAM_OBJ_Pose= visor_getPose3d (1, 0)
          $ 1286 "If CAM_CNT_Obj>0"
          if (CAM_CNT_Obj>0):
            $ 1287 "CAM_OBJ_Color≔visor_getAdditionalData(1, 0)"
            global CAM_OBJ_Color= visor_getAdditionalData (1, 0)
            $ 1288 "CAM_DetectScore≔to_num(visor_getAdditionalData(1, 1))/1000"
            global CAM_DetectScore=to_num( visor_getAdditionalData (1, 1))/1000
            $ 1289 "OBJ_Detected≔ True "
            global OBJ_Detected=  True
          end
        else:
          $ 1290 "Else" "noBreak"
          $ 1291 "CAM_Captures≔CAM_Captures+1"
          global CAM_Captures=CAM_Captures+1
        end
        $ 1292 "If OBJ_Detected"
        if (OBJ_Detected):
          $ 1293 "Get object data"
          $ 1294 "PRC_CntDetect≔0"
          global PRC_CntDetect=0
          $ 1295 "Loop PRC_CntDetect<CAM_CNT_Obj"
          while (PRC_CntDetect<CAM_CNT_Obj):
            $ 1296 "get object and jig number"
            $ 1297 "If ITM_ID≟1 and JIG≟7"
            if (ITM_ID == 1  and  JIG == 7):
              $ 1298 "FRM_Reference≔FRM_Cap_SSRack"
              global FRM_Reference=FRM_Cap_SSRack
            else:
              $ 1299 "ElseIf ITM_ID≟5 and JIG≟7"
              if (ITM_ID == 5  and  JIG == 7):
                $ 1300 "FRM_Reference≔uLM_Cap_SSRack"
                global FRM_Reference=uLM_Cap_SSRack
              end
            end
            $ 1303 "PSE_T≔pose_trans(pose_inv(FRM_Reference), CAM_OBJ_Pose)"
            global PSE_T= pose_trans ( pose_inv (FRM_Reference), CAM_OBJ_Pose)
            $ 1304 "CAM_Result.append(get_pattern_counter(PSE_T, 'X', pattern=[10, 5], patternsize=[0.181, 0.081]))"
            CAM_Result.append(get_pattern_counter(PSE_T, "X", pattern=[10, 5], patternsize=[0.181, 0.081]))
            $ 1305 "PRC_CntDetect≔PRC_CntDetect+1"
            global PRC_CntDetect=PRC_CntDetect+1
          end
          $ 1306 "CAM_Done≔ True "
          global CAM_Done=  True
        else:
          $ 1307 "ElseIf CAM_Captures≥CAM_PRM_Retries"
          if (CAM_Captures >= CAM_PRM_Retries):
            $ 1308 "CAM_Done≔ True "
            global CAM_Done=  True
          else:
            $ 1309 "Else" "noBreak"
            $ 1310 "CAM_Captures≔CAM_Captures+1"
            global CAM_Captures=CAM_Captures+1
          end
        end
      end
    end
    $ 1311 "'=========='"
    # '=========='
    $ 1312 "PostSettings"
    $ 1313 "FRM_Reference≔p[0,0,0,0,0,0]"
    global FRM_Reference=p[0,0,0,0,0,0]
    $ 1314 "Set"
    set_tcp(p[0.0,0.0,0.161,3.1415,0.0,0.0])
    $ 1315 "CAM_Pose≔p[0,0,0,0,0,0]"
    global CAM_Pose=p[0,0,0,0,0,0]
    $ 1316 "Action≔0"
    global Action=0
    $ 1317 "Action_Info≔''"
    global Action_Info=""
  end
  def Sub_AMR_MiR_V3():
    $ 1318 "Sub_AMR_MiR_V3" "noBreak"
    $ 1319 "PreSettings"
    $ 1320 "AMR_TargetList≔[1,2,3,4,5,6,7,21,22,23,24,31,32,33,34,35,36,37,38,41]"
    global AMR_TargetList=[1,2,3,4,5,6,7,21,22,23,24,31,32,33,34,35,36,37,38,41]
    $ 1321 "AMR_Done≔ False "
    global AMR_Done=  False
    $ 1322 "AMR_PosActual≔T2O_Current_Pos"
    global AMR_PosActual=modbus_get_signal_status("T2O_Current_Pos")
    $ 1323 "AMR_Attemps≔T2O_Nav_Attemps"
    global AMR_Attemps=modbus_get_signal_status("T2O_Nav_Attemps")
    $ 1324 "AMR_Battery≔MiR_Battery_Lvl"
    global AMR_Battery=modbus_get_signal_status("MiR_Battery_Lvl")
    $ 1325 "AMR_Charging≔(T2O_Charging≟1)"
    global AMR_Charging=(modbus_get_signal_status("T2O_Charging") == 1)
    $ 1326 "AMR_Position≔struct(position_identifier=T2O_Current_Pos, x1=MiR_Position_X1, x2=MiR_Position_X2, y1=MiR_Position_Y1, y2=MiR_Position_Y2, theta1=MiR_Theta_1, theta2=MiR_Theta_2) "
    global AMR_Position=struct(position_identifier=modbus_get_signal_status("T2O_Current_Pos"), x1=modbus_get_signal_status("MiR_Position_X1"), x2=modbus_get_signal_status("MiR_Position_X2"), y1=modbus_get_signal_status("MiR_Position_Y1"), y2=modbus_get_signal_status("MiR_Position_Y2"), theta1=modbus_get_signal_status("MiR_Theta_1"), theta2=modbus_get_signal_status("MiR_Theta_2"))
    $ 1327 "If MiR_Mode≠7"
    if (modbus_get_signal_status("MiR_Mode") != 7):
      $ 1328 "Error"
      $ 1329 "set_error(ERROR_AMR_WRONG_MODE)"
      set_error(ERROR_AMR_WRONG_MODE)
      $ 1330 "AMR_Done≔ True "
      global AMR_Done=  True
    end
    $ 1331 "'=========='"
    # '=========='
    $ 1332 "Switch STATE"
    switch_1 = STATE
    $ 1333 "Case 1"
    if (1 == switch_1):
      $ 1334 "stopping"
      $ 1335 "If T2O_Done≟1 and O2T_Acknowledge≟0"
      if (modbus_get_signal_status("T2O_Done") == 1  and  modbus_get_signal_status("O2T_Acknowledge") == 0):
        $ 1336 "Set O2T_Acknowledge=1"
        modbus_set_output_register("O2T_Acknowledge", 1)
      end
      $ 1337 "Set MiR_CMD_Stop=On"
      modbus_set_output_signal("MiR_CMD_Stop", True)
      $ 1338 "AMR_Position.position_identifier = 0"
      AMR_Position.position_identifier = 0
      $ 1339 "AMR_Done≔ True "
      global AMR_Done=  True
    elif (2 == switch_1):
      $ 1340 "Case 2"
      $ 1341 "stopped"
      $ 1342 "If MiR_State≠3 and MiR_State≠5"
      if (modbus_get_signal_status("MiR_State") != 3  and  modbus_get_signal_status("MiR_State") != 5):
        $ 1343 "Set MiR_CMD_Stop=Off"
        modbus_set_output_signal("MiR_CMD_Stop", False)
      end
    elif (3 == switch_1):
      $ 1344 "Case 3"
      $ 1345 "resetting"
      $ 1346 "Set O2T_Mis_Main=Off"
      modbus_set_output_signal("O2T_Mis_Main", False)
      $ 1347 "Set O2T_Mis_Charge=Off"
      modbus_set_output_signal("O2T_Mis_Charge", False)
      $ 1348 "If MiR_Mis_Queue>0"
      if (modbus_get_signal_status("MiR_Mis_Queue")>0):
        $ 1349 "Set MiR_CMD_Clear_Q=On"
        modbus_set_output_signal("MiR_CMD_Clear_Q", True)
        $ 1350 "Wait MiR_Mis_Queue≟0"
        while (not(modbus_get_signal_status("MiR_Mis_Queue") == 0)):
          sync()
        end
        $ 1351 "Set MiR_CMD_Clear_Q=Off"
        modbus_set_output_signal("MiR_CMD_Clear_Q", False)
      end
      $ 1352 "If MiR_Error_ID≠0"
      if (modbus_get_signal_status("MiR_Error_ID") != 0):
        $ 1353 "Set MiR_CMD_Clear_E=On"
        modbus_set_output_signal("MiR_CMD_Clear_E", True)
        $ 1354 "Wait MiR_Error_ID≟0"
        while (not(modbus_get_signal_status("MiR_Error_ID") == 0)):
          sync()
        end
        $ 1355 "Set MiR_CMD_Clear_E=Off"
        modbus_set_output_signal("MiR_CMD_Clear_E", False)
      end
      $ 1356 "Set O2T_Action=0"
      modbus_set_output_register("O2T_Action", 0)
      $ 1357 "Set O2T_Acknowledge=0"
      modbus_set_output_register("O2T_Acknowledge", 0)
      $ 1358 "Set O2T_Target_Pos=0"
      modbus_set_output_register("O2T_Target_Pos", 0)
      $ 1359 "Set O2T_Footprint=0"
      modbus_set_output_register("O2T_Footprint", 0)
      $ 1360 "Set O2T_ProtectOff=0"
      modbus_set_output_register("O2T_ProtectOff", 0)
      $ 1361 "Set O2T_Dock=0"
      modbus_set_output_register("O2T_Dock", 0)
      $ 1362 "AMR_Attemps≔0"
      global AMR_Attemps=0
      $ 1363 "AMR_PosTarget≔0"
      global AMR_PosTarget=0
      $ 1364 "AMR_Step≔0"
      global AMR_Step=0
      $ 1365 "AMR_AtTarget≔ False "
      global AMR_AtTarget=  False
      $ 1366 "If MiR_State≟4 or MiR_State≟3 or MiR_State≟10"
      if (modbus_get_signal_status("MiR_State") == 4  or  modbus_get_signal_status("MiR_State") == 3  or  modbus_get_signal_status("MiR_State") == 10):
        $ 1367 "AMR_Done≔ True "
        global AMR_Done=  True
      end
    elif (5 == switch_1):
      $ 1368 "Case 5"
      $ 1369 "starting"
      $ 1370 "If MiR_State≟4"
      if (modbus_get_signal_status("MiR_State") == 4):
        $ 1371 "Set MiR_CMD_Start=On"
        modbus_set_output_signal("MiR_CMD_Start", True)
        $ 1372 "Wait MiR_State≠4"
        while (not(modbus_get_signal_status("MiR_State") != 4)):
          sync()
        end
        $ 1373 "Set MiR_CMD_Start=Off"
        modbus_set_output_signal("MiR_CMD_Start", False)
        $ 1374 "AMR_Done≔ True "
        global AMR_Done=  True
      else:
        $ 1375 "ElseIf MiR_State≟10"
        if (modbus_get_signal_status("MiR_State") == 10):
          $ 1376 "'MiR in protective stop. Wait'"
          # 'MiR in protective stop. Wait'
          $ 1377 "AMR_Done≔ True "
          global AMR_Done=  True
        else:
          $ 1378 "ElseIf MiR_State≟3"
          if (modbus_get_signal_status("MiR_State") == 3):
            $ 1379 "AMR_Done≔ True "
            global AMR_Done=  True
          end
        end
      end
    elif (6 == switch_1):
      $ 1380 "Case 6"
      $ 1381 "execute"
      $ 1382 "AMR_AtTarget≔(AMR_PosActual≟AMR_PosTarget)"
      global AMR_AtTarget=(AMR_PosActual == AMR_PosTarget)
      $ 1383 "Switch AMR_Step"
      switch_2 = AMR_Step
      $ 1384 "Case 0"
      if (0 == switch_2):
        $ 1385 "If  not AMR_AtTarget"
        if (  not  AMR_AtTarget):
          $ 1386 "AMR_Step≔1"
          global AMR_Step=1
        else:
          $ 1387 "Else" "noBreak"
          $ 1388 "AMR_Done≔ True "
          global AMR_Done=  True
        end
      elif (1 == switch_2):
        $ 1389 "Case 1"
        $ 1390 "general Settings"
        $ 1391 "Set O2T_Acknowledge=0"
        modbus_set_output_register("O2T_Acknowledge", 0)
        $ 1392 "check for error"
        $ 1393 "If OBJ_Picked and MiR_State≟10"
        if (OBJ_Picked  and  modbus_get_signal_status("MiR_State") == 10):
          $ 1394 "Error"
          $ 1395 "set_error(ERROR_ROBOT_ARM_NOT_IN_HOME_POSE)"
          set_error(ERROR_ROBOT_ARM_NOT_IN_HOME_POSE)
          $ 1396 "Action≔0"
          global Action=0
        else:
          $ 1397 "ElseIf  not found_in_list(AMR_PosTarget, AMR_TargetList)"
          if (  not  found_in_list(AMR_PosTarget, AMR_TargetList)):
            $ 1398 "Error"
            $ 1399 "set_error(ERROR_UNKNOWN_POSE)"
            set_error(ERROR_UNKNOWN_POSE)
            $ 1400 "Action≔0"
            global Action=0
          end
        end
        $ 1401 "If MiR_State≟3"
        if (modbus_get_signal_status("MiR_State") == 3):
          $ 1402 "Set MiR_CMD_Start=Off"
          modbus_set_output_signal("MiR_CMD_Start", False)
          $ 1403 "Switch Action"
          switch_3 = Action
          $ 1404 "Case 51"
          if (51 == switch_3):
            $ 1405 "Charge"
            $ 1406 "'trigger the charging mission'"
            # 'trigger the charging mission'
            $ 1407 "'target pos is predefined'"
            # 'target pos is predefined'
            $ 1408 "Set O2T_Footprint=0"
            modbus_set_output_register("O2T_Footprint", 0)
            $ 1409 "Set O2T_Action=1"
            modbus_set_output_register("O2T_Action", 1)
            $ 1410 "If MiR_Mis_Queue≟0"
            if (modbus_get_signal_status("MiR_Mis_Queue") == 0):
              $ 1411 "Set O2T_Mis_Charge=On"
              modbus_set_output_signal("O2T_Mis_Charge", True)
              $ 1412 "Wait MiR_Mis_Queue≥1"
              while (not(modbus_get_signal_status("MiR_Mis_Queue") >= 1)):
                sync()
              end
              $ 1413 "Set O2T_Mis_Charge=Off"
              modbus_set_output_signal("O2T_Mis_Charge", False)
            end
          elif (52 == switch_3):
            $ 1414 "Case 52"
            $ 1415 "Navigate"
            $ 1416 "'trigger the standard missoin'"
            # 'trigger the standard missoin'
            $ 1417 "Set O2T_Footprint=AMR_FootprintID"
            modbus_set_output_register("O2T_Footprint", AMR_FootprintID)
            $ 1418 "Set O2T_Target_Pos=AMR_PosTarget"
            modbus_set_output_register("O2T_Target_Pos", AMR_PosTarget)
            $ 1419 "Set O2T_Action=2"
            modbus_set_output_register("O2T_Action", 2)
            $ 1420 "If MiR_Mis_Queue≟0"
            if (modbus_get_signal_status("MiR_Mis_Queue") == 0):
              $ 1421 "Set O2T_Mis_Main=On"
              modbus_set_output_signal("O2T_Mis_Main", True)
              $ 1422 "Wait MiR_Mis_Queue≥1"
              while (not(modbus_get_signal_status("MiR_Mis_Queue") >= 1)):
                sync()
              end
              $ 1423 "Set O2T_Mis_Main=Off"
              modbus_set_output_signal("O2T_Mis_Main", False)
            end
          end
        else:
          $ 1424 "ElseIf MiR_State≟4"
          if (modbus_get_signal_status("MiR_State") == 4):
            $ 1425 "Set MiR_CMD_Start=On"
            modbus_set_output_signal("MiR_CMD_Start", True)
          else:
            $ 1426 "ElseIf MiR_State≟5"
            if (modbus_get_signal_status("MiR_State") == 5):
              $ 1427 "AMR_Step≔2"
              global AMR_Step=2
            else:
              $ 1428 "ElseIf MiR_State≟10"
              if (modbus_get_signal_status("MiR_State") == 10):
                $ 1429 "'AMR still in safeguard stop'"
                # 'AMR still in safeguard stop'
              end
            end
          end
        end
      elif (2 == switch_2):
        $ 1430 "Case 2"
        $ 1431 "acknowledge handshake"
        $ 1432 "If T2O_Done≟1 and O2T_Acknowledge≟0"
        if (modbus_get_signal_status("T2O_Done") == 1  and  modbus_get_signal_status("O2T_Acknowledge") == 0):
          $ 1433 "Set O2T_Acknowledge=1"
          modbus_set_output_register("O2T_Acknowledge", 1)
        else:
          $ 1434 "ElseIf T2O_Done≟0 and O2T_Acknowledge≟1"
          if (modbus_get_signal_status("T2O_Done") == 0  and  modbus_get_signal_status("O2T_Acknowledge") == 1):
            $ 1435 "Set O2T_Acknowledge=0"
            modbus_set_output_register("O2T_Acknowledge", 0)
            $ 1436 "AMR_AtTarget≔(AMR_PosActual≟AMR_PosTarget)"
            global AMR_AtTarget=(AMR_PosActual == AMR_PosTarget)
            $ 1437 "AMR_Done≔ True "
            global AMR_Done=  True
          end
        end
      end
      $ 1438 "translate errors"
      $ 1439 "If AMR_Done"
      if (AMR_Done):
        $ 1440 "Switch T2O_Error_ID"
        switch_2 = modbus_get_signal_status("T2O_Error_ID")
        $ 1441 "Case 2003"
        if (2003 == switch_2):
          $ 1442 "error"
          $ 1443 "set_error(ERROR_NOT_DOCKED)"
          set_error(ERROR_NOT_DOCKED)
        elif (2007 == switch_2):
          $ 1444 "Case 2007"
          $ 1445 "error"
          $ 1446 "set_error(ERROR_NOT_REACHABLE_TARGET)"
          set_error(ERROR_NOT_REACHABLE_TARGET)
        elif (2008 == switch_2):
          $ 1447 "Case 2008"
          $ 1448 "error"
          $ 1449 "set_error(ERROR_CHARGING_NOT_STARTED)"
          set_error(ERROR_CHARGING_NOT_STARTED)
        end
      end
    elif (7 == switch_1):
      $ 1450 "Case 7"
      $ 1451 "completing"
      $ 1452 "If MiR_Mis_Queue>0"
      if (modbus_get_signal_status("MiR_Mis_Queue")>0):
        $ 1453 "Set MiR_CMD_Abort=On"
        modbus_set_output_signal("MiR_CMD_Abort", True)
        $ 1454 "Wait MiR_Mis_Queue≟0"
        while (not(modbus_get_signal_status("MiR_Mis_Queue") == 0)):
          sync()
        end
        $ 1455 "Set MiR_CMD_Abort=Off"
        modbus_set_output_signal("MiR_CMD_Abort", False)
      end
      $ 1456 "If MiR_State≟3 or MiR_State≟10"
      if (modbus_get_signal_status("MiR_State") == 3  or  modbus_get_signal_status("MiR_State") == 10):
        $ 1457 "AMR_Done≔ True "
        global AMR_Done=  True
      end
    elif (9 == switch_1):
      $ 1458 "Case 9"
      $ 1459 "holding"
      $ 1460 "Set MiR_CMD_Abort=On"
      modbus_set_output_signal("MiR_CMD_Abort", True)
      $ 1461 "If MiR_State≟3 or MiR_State≟10"
      if (modbus_get_signal_status("MiR_State") == 3  or  modbus_get_signal_status("MiR_State") == 10):
        $ 1462 "Set MiR_CMD_Abort=Off"
        modbus_set_output_signal("MiR_CMD_Abort", False)
        $ 1463 "AMR_Done≔ True "
        global AMR_Done=  True
      end
    elif (11 == switch_1):
      $ 1464 "Case 11"
      $ 1465 "unholding"
      $ 1466 "Set MiR_CMD_Start=On"
      modbus_set_output_signal("MiR_CMD_Start", True)
      $ 1467 "If MiR_State≠4"
      if (modbus_get_signal_status("MiR_State") != 4):
        $ 1468 "Set MiR_CMD_Start=Off"
        modbus_set_output_signal("MiR_CMD_Start", False)
        $ 1469 "AMR_Step≔0"
        global AMR_Step=0
        $ 1470 "AMR_Done≔ True "
        global AMR_Done=  True
      end
    elif (12 == switch_1):
      $ 1471 "Case 12"
      $ 1472 "suspending"
      $ 1473 "'none'"
      # 'none'
    elif (14 == switch_1):
      $ 1474 "Case 14"
      $ 1475 "unsuspending"
      $ 1476 "'none'"
      # 'none'
    elif (15 == switch_1):
      $ 1477 "Case 15"
      $ 1478 "aborting"
      $ 1479 "Set MiR_CMD_Abort=On"
      modbus_set_output_signal("MiR_CMD_Abort", True)
      $ 1480 "Wait MiR_State≟3"
      while (not(modbus_get_signal_status("MiR_State") == 3)):
        sync()
      end
      $ 1481 "Set MiR_CMD_Abort=Off"
      modbus_set_output_signal("MiR_CMD_Abort", False)
    elif (17 == switch_1):
      $ 1482 "Case 17"
      $ 1483 "clearing"
      $ 1484 "If MiR_Error_ID≠0"
      if (modbus_get_signal_status("MiR_Error_ID") != 0):
        $ 1485 "Set MiR_CMD_Clear_E=On"
        modbus_set_output_signal("MiR_CMD_Clear_E", True)
        $ 1486 "Wait MiR_Error_ID≟0"
        while (not(modbus_get_signal_status("MiR_Error_ID") == 0)):
          sync()
        end
        $ 1487 "Set MiR_CMD_Clear_E=Off"
        modbus_set_output_signal("MiR_CMD_Clear_E", False)
      end
      $ 1488 "If MiR_Error_ID≟0"
      if (modbus_get_signal_status("MiR_Error_ID") == 0):
        $ 1489 "AMR_Done≔ True "
        global AMR_Done=  True
      end
    end
    $ 1490 "'=========='"
    # '=========='
    $ 1491 "PostSettings"
    $ 1492 "AMR_Position≔struct(position_identifier=T2O_Current_Pos, x1=MiR_Position_X1, x2=MiR_Position_X2, y1=MiR_Position_Y1, y2=MiR_Position_Y2, theta1=MiR_Theta_1, theta2=MiR_Theta_2) "
    global AMR_Position=struct(position_identifier=modbus_get_signal_status("T2O_Current_Pos"), x1=modbus_get_signal_status("MiR_Position_X1"), x2=modbus_get_signal_status("MiR_Position_X2"), y1=modbus_get_signal_status("MiR_Position_Y1"), y2=modbus_get_signal_status("MiR_Position_Y2"), theta1=modbus_get_signal_status("MiR_Theta_1"), theta2=modbus_get_signal_status("MiR_Theta_2"))
  end
  def Sub_Action_V4():
    $ 1493 "Sub_Action_V4" "noBreak"
    $ 1494 "PreSettings"
    $ 1495 "init poses"
    $ 1496 "PSE_A≔p[0,0,0,0,0,0]"
    global PSE_A=p[0,0,0,0,0,0]
    $ 1497 "PSE_A_H≔p[0,0,0,0,0,0]"
    global PSE_A_H=p[0,0,0,0,0,0]
    $ 1498 "PSE_T≔p[0,0,0,0,0,0]"
    global PSE_T=p[0,0,0,0,0,0]
    $ 1499 "PSE_T_H≔p[0,0,0,0,0,0]"
    global PSE_T_H=p[0,0,0,0,0,0]
    $ 1500 "PSE_G≔p[0,0,0,0,0,0]"
    global PSE_G=p[0,0,0,0,0,0]
    $ 1501 "PSE_G_H≔p[0,0,0,0,0,0]"
    global PSE_G_H=p[0,0,0,0,0,0]
    $ 1502 "PSE_R≔p[0,0,0,0,0,0]"
    global PSE_R=p[0,0,0,0,0,0]
    $ 1503 "PSE_R_H≔p[0,0,0,0,0,0]"
    global PSE_R_H=p[0,0,0,0,0,0]
    $ 1504 "JNT_Q≔[0,0,0,0,0,0]"
    global JNT_Q=[0,0,0,0,0,0]
    $ 1505 "JNT_S≔[0,0,0,0,0,0]"
    global JNT_S=[0,0,0,0,0,0]
    $ 1506 "Gripping parameters"
    $ 1507 "OBJ = find_object_by_type(OBJs, OBJ_Type)"
    OBJ = find_object_by_type(OBJs, OBJ_Type)
    $ 1508 "GRP_Open_Pos≔OBJ.dimension.diameter * 1000 + 6"
    global GRP_Open_Pos=OBJ.dimension.diameter * 1000 + 6
    $ 1509 "GRP_Offset≔OBJ.gripper_offset"
    global GRP_Offset=OBJ.gripper_offset
    $ 1510 "rq_set_force_norm(50)"
     rq_set_force_norm (50)
    $ 1511 "rq_set_speed_norm(50)"
     rq_set_speed_norm (50)
    $ 1512 "Switch ITM_ID"
    switch_1 = ITM_ID
    $ 1513 "Case 1"
    if (1 == switch_1):
      $ 1514 "uML"
      $ 1515 "JIG2 = find_object_by_type(JIGs, JIG)"
      JIG2 = find_object_by_type(JIGs, JIG)
      $ 1516 "JIG_Offset≔JIG2.jig_offset"
      global JIG_Offset=JIG2.jig_offset
      $ 1517 "Switch JIG"
      switch_2 = JIG
      $ 1518 "Case 1"
      if (1 == switch_2):
        $ 1519 "3FG"
        $ 1520 "define poses"
        $ 1521 "FRM_Reference≔ULM_3FG"
        global FRM_Reference=ULM_3FG
        $ 1522 "JNT_Q≔JNT_HOME"
        global JNT_Q=JNT_HOME
        $ 1523 "PSE_T≔pose_trans(GRP_Offset, JIG_Offset)"
        global PSE_T= pose_trans (GRP_Offset, JIG_Offset)
        $ 1524 "PSE_A≔pose_trans(PSE_T, p[0,0,0.100,0,0,0])"
        global PSE_A= pose_trans (PSE_T, p[0,0,0.100,0,0,0])
        $ 1525 "PSE_R≔pose_add(PSE_T, p[0,0,0.100,0,0,0])"
        global PSE_R= pose_add (PSE_T, p[0,0,0.100,0,0,0])
      elif (2 == switch_2):
        $ 1526 "Case 2"
        $ 1527 "Input"
        $ 1528 "'CHANGE THE REFERENCE TO THE FRAME TO MOVE IN'"
        # 'CHANGE THE REFERENCE TO THE FRAME TO MOVE IN'
        $ 1529 "define poses"
        $ 1530 "FRM_Reference≔ULM_Input"
        global FRM_Reference=ULM_Input
        $ 1531 "PSE_T≔pose_trans(pose_trans(get_pattern_pos_rectangle(OBJ_Nbr, 'X', [10,5], patternsize=[0.181,0.081]), GRP_Offset), JIG_Offset)"
        global PSE_T= pose_trans ( pose_trans (get_pattern_pos_rectangle(OBJ_Nbr, "X", [10,5], patternsize=[0.181,0.081]), GRP_Offset), JIG_Offset)
        $ 1532 "If Action≟1"
        if (Action == 1):
          $ 1533 "PSE_R≔pose_add(PSE_T, p[0,0,0.200,0,0,0])"
          global PSE_R= pose_add (PSE_T, p[0,0,0.200,0,0,0])
          $ 1534 "PSE_A≔pose_add(PSE_T, p[0,0,0.100,0,0,0])"
          global PSE_A= pose_add (PSE_T, p[0,0,0.100,0,0,0])
        else:
          $ 1535 "ElseIf Action≟2"
          if (Action == 2):
            $ 1536 "PSE_R≔pose_add(PSE_T, p[0,0,0.100,0,0,0])"
            global PSE_R= pose_add (PSE_T, p[0,0,0.100,0,0,0])
            $ 1537 "PSE_A≔pose_add(PSE_T, p[0,0,0.200,0,0,0])"
            global PSE_A= pose_add (PSE_T, p[0,0,0.200,0,0,0])
          end
        end
      elif (3 == switch_2):
        $ 1538 "Case 3"
        $ 1539 "Output"
        $ 1540 "'CHANGE THE REFERENCE TO THE FRAME TO MOVE IN'"
        # 'CHANGE THE REFERENCE TO THE FRAME TO MOVE IN'
        $ 1541 "define poses"
        $ 1542 "FRM_Reference≔ULM_Output"
        global FRM_Reference=ULM_Output
        $ 1543 "PSE_T≔pose_trans(pose_trans(get_pattern_pos_rectangle(OBJ_Nbr, 'X', [10,5], patternsize=[0.181,0.081]), GRP_Offset), JIG_Offset)"
        global PSE_T= pose_trans ( pose_trans (get_pattern_pos_rectangle(OBJ_Nbr, "X", [10,5], patternsize=[0.181,0.081]), GRP_Offset), JIG_Offset)
        $ 1545 "If Action≟1"
        if (Action == 1):
          $ 1546 "PSE_R≔pose_add(PSE_T, p[0,0,0.200,0,0,0])"
          global PSE_R= pose_add (PSE_T, p[0,0,0.200,0,0,0])
          $ 1547 "PSE_A≔pose_add(PSE_T, p[0,0,0.100,0,0,0])"
          global PSE_A= pose_add (PSE_T, p[0,0,0.100,0,0,0])
        else:
          $ 1548 "ElseIf Action≟2"
          if (Action == 2):
            $ 1549 "PSE_R≔pose_add(PSE_T, p[0,0,0.100,0,0,0])"
            global PSE_R= pose_add (PSE_T, p[0,0,0.100,0,0,0])
            $ 1550 "PSE_A≔pose_add(PSE_T, p[0,0,0.200,0,0,0])"
            global PSE_A= pose_add (PSE_T, p[0,0,0.200,0,0,0])
          end
        end
      elif (4 == switch_2):
        $ 1551 "Case 4"
        $ 1552 "jig centrifuge racks"
        $ 1553 "define poses"
        $ 1554 "FRM_Reference≔ULM_Cent_Racks"
        global FRM_Reference=ULM_Cent_Racks
        $ 1555 "PSE_T≔get_pattern_pos_rectangle(JIG_Slot, 'X', [4,1], patternsize=[0.291,0])"
        global PSE_T=get_pattern_pos_rectangle(JIG_Slot, "X", [4,1], patternsize=[0.291,0])
        $ 1556 "If OBJ_Nbr≠0"
        if (OBJ_Nbr != 0):
          $ 1557 "PSE_T≔pose_trans(pose_trans(PSE_T, get_pattern_pos_rectangle(OBJ_Nbr, 'X', [3,3], patternsize=[0.060,0.060])),p[-0.030, -0.030,0,0,0,3.927])"
          global PSE_T= pose_trans ( pose_trans (PSE_T, get_pattern_pos_rectangle(OBJ_Nbr, "X", [3,3], patternsize=[0.060,0.060])),p[-0.030, -0.030,0,0,0,3.927])
        end
        $ 1558 "PSE_T≔pose_trans(PSE_T, GRP_Offset)"
        global PSE_T= pose_trans (PSE_T, GRP_Offset)
        $ 1559 "If Action≟1"
        if (Action == 1):
          $ 1560 "PSE_R≔pose_add(PSE_T, p[0,0,0.200,0,0,0])"
          global PSE_R= pose_add (PSE_T, p[0,0,0.200,0,0,0])
          $ 1561 "PSE_A≔pose_add(PSE_T, p[0,0,0.100,0,0,0])"
          global PSE_A= pose_add (PSE_T, p[0,0,0.100,0,0,0])
        else:
          $ 1562 "ElseIf Action≟2"
          if (Action == 2):
            $ 1563 "PSE_R≔pose_add(PSE_T, p[0,0,0.100,0,0,0])"
            global PSE_R= pose_add (PSE_T, p[0,0,0.100,0,0,0])
            $ 1564 "PSE_A≔pose_add(PSE_T, p[0,0,0.200,0,0,0])"
            global PSE_A= pose_add (PSE_T, p[0,0,0.200,0,0,0])
          end
        end
      elif (6 == switch_2):
        $ 1565 "Case 6"
        $ 1566 "Caps bin"
        $ 1567 "define poses"
        $ 1568 "'Drop cap'"
        # 'Drop cap'
        $ 1569 "FRM_Reference=ULM_Cap_Bin"
        FRM_Reference=ULM_Cap_Bin
        $ 1570 "PSE_T≔pose_RPY2RotVec(p[0,0,0,0,0,0])"
        global PSE_T=pose_RPY2RotVec(p[0,0,0,0,0,0])
        $ 1571 "PSE_T_H≔pose_add(PSE_T, p[0,0,-0.011,0,0,0])"
        global PSE_T_H= pose_add (PSE_T, p[0,0,-0.011,0,0,0])
        $ 1572 "PSE_A≔pose_trans(PSE_T, p[0,0,0.1,0,0,0])"
        global PSE_A= pose_trans (PSE_T, p[0,0,0.1,0,0,0])
        $ 1573 "PSE_R_H≔pose_add(PSE_T, p[0,0,0.100,0,0,0])"
        global PSE_R_H= pose_add (PSE_T, p[0,0,0.100,0,0,0])
        $ 1574 "PSE_R≔pose_add(PSE_T, p[0,0,0.100,0,0,0])"
        global PSE_R= pose_add (PSE_T, p[0,0,0.100,0,0,0])
      elif (7 == switch_2):
        $ 1575 "Case 7"
      elif (8 == switch_2):
        $ 1600 "Case 8"
        $ 1601 "NoK"
        $ 1602 "define poses"
        $ 1603 "'NoK'"
        # 'NoK'
        $ 1604 "FRM_Reference=ULM_NoK"
        FRM_Reference=ULM_NoK
        $ 1605 "PSE_T≔pose_RPY2RotVec(p[0,0,0,0,0,0])"
        global PSE_T=pose_RPY2RotVec(p[0,0,0,0,0,0])
        $ 1606 "PSE_A≔pose_trans(PSE_T, p[0,0,0.1,0,0,0])"
        global PSE_A= pose_trans (PSE_T, p[0,0,0.1,0,0,0])
        $ 1607 "PSE_R≔pose_add(PSE_T, p[0,0,0.100,0,0,0])"
        global PSE_R= pose_add (PSE_T, p[0,0,0.100,0,0,0])
      elif (9 == switch_2):
        $ 1608 "Case 9"
      elif (10 == switch_2):
        $ 1616 "Case 10"
      elif (11 == switch_2):
        $ 1624 "Case 11"
      elif (12 == switch_2):
        $ 1632 "Case 12"
      end
    elif (2 == switch_1):
      $ 1640 "Case 2"
      $ 1641 "Centrifuge"
      $ 1642 "'CHANGE THE REFERENCE TO THE FRAME TO MOVE IN'"
      # 'CHANGE THE REFERENCE TO THE FRAME TO MOVE IN'
      $ 1643 "define poses"
      $ 1644 "FRM_Reference≔FRM_Centrifuge"
      global FRM_Reference=FRM_Centrifuge
      $ 1645 "PSE_T≔GRP_Offset"
      global PSE_T=GRP_Offset
      $ 1646 "If Action≟8"
      if (Action == 8):
        $ 1647 "PSE_R≔pose_add(PSE_T, p[0,0,0.250,0,0,0])"
        global PSE_R= pose_add (PSE_T, p[0,0,0.250,0,0,0])
        $ 1648 "PSE_A≔pose_add(PSE_T, p[0,0,0.150,0,0,0])"
        global PSE_A= pose_add (PSE_T, p[0,0,0.150,0,0,0])
      else:
        $ 1649 "ElseIf Action≟7"
        if (Action == 7):
          $ 1650 "PSE_R≔pose_add(PSE_T, p[0,0,0.150,0,0,0])"
          global PSE_R= pose_add (PSE_T, p[0,0,0.150,0,0,0])
          $ 1651 "PSE_A≔pose_add(PSE_T, p[0,0,0.250,0,0,0])"
          global PSE_A= pose_add (PSE_T, p[0,0,0.250,0,0,0])
        end
      end
    elif (3 == switch_1):
      $ 1652 "Case 3"
      $ 1653 "Output"
      $ 1654 "'CHANGE THE REFERENCE TO THE FRAME TO MOVE IN'"
      # 'CHANGE THE REFERENCE TO THE FRAME TO MOVE IN'
      $ 1655 "define poses"
      $ 1656 "FRM_Reference≔Base_const"
      global FRM_Reference=p[0.0,0.0,0.0,0.0,0.0,0.0]
      $ 1657 "PSE_T≔p[0,0,0,0,0,0]"
      global PSE_T=p[0,0,0,0,0,0]
      $ 1658 "PSE_A≔pose_add(PSE_T, p[0,0,0.150,0,0,0])"
      global PSE_A= pose_add (PSE_T, p[0,0,0.150,0,0,0])
      $ 1659 "PSE_R≔pose_add(PSE_T, p[0,0,0.100,0,0,0])"
      global PSE_R= pose_add (PSE_T, p[0,0,0.100,0,0,0])
    elif (5 == switch_1):
      $ 1660 "Case 5"
      $ 1661 "Sarstedt Pickup Table"
      $ 1662 "'CHANGE THE REFERENCE TO THE FRAME TO MOVE IN'"
      # 'CHANGE THE REFERENCE TO THE FRAME TO MOVE IN'
      $ 1663 "Switch JIG"
      switch_2 = JIG
      $ 1664 "Case 7"
      if (7 == switch_2):
        $ 1677 "Sarstedt"
        $ 1678 "'CHANGE THE REFERENCE TO THE FRAME TO MOVE IN'"
        # 'CHANGE THE REFERENCE TO THE FRAME TO MOVE IN'
        $ 1684 "If TASK.ID≟10"
        if (TASK.ID == 10):
          $ 1685 "Frame & Position Params"
          $ 1686 "FRM_Reference = CAM_LM_SSRack"
          FRM_Reference = CAM_LM_SSRack
          $ 1687 "PSE_T≔uLM_SS_PickPlc"
          global PSE_T=uLM_SS_PickPlc
          $ 1688 "PSE_A≔pose_trans(PSE_T, p[0,0,0.1,0,0,0])"
          global PSE_A= pose_trans (PSE_T, p[0,0,0.1,0,0,0])
          $ 1689 "PSE_R≔pose_add(PSE_T, p[0,0,0.1,0,0,0])"
          global PSE_R= pose_add (PSE_T, p[0,0,0.1,0,0,0])
        end
      end
    elif (13 == switch_1):
      $ 1696 "Case 13"
      $ 1697 "Sarstedt Pickup Table"
      $ 1698 "'CHANGE THE REFERENCE TO THE FRAME TO MOVE IN'"
      # 'CHANGE THE REFERENCE TO THE FRAME TO MOVE IN'
      $ 1699 "Switch JIG"
      switch_2 = JIG
      $ 1700 "Case 7"
      if (7 == switch_2):
        $ 1713 "Bottle"
        $ 1714 "'CHANGE THE REFERENCE TO THE FRAME TO MOVE IN'"
        # 'CHANGE THE REFERENCE TO THE FRAME TO MOVE IN'
        $ 1720 "If TASK.ID≟43"
        if (TASK.ID == 43):
          $ 1721 "Frame & Position Params"
          $ 1723 "PSE_T≔uLM_SS_PickPlc"
          global PSE_T=uLM_SS_PickPlc
          $ 1724 "PSE_A≔pose_trans(PSE_T, p[0,0,0.1,0,0,0])"
          global PSE_A= pose_trans (PSE_T, p[0,0,0.1,0,0,0])
          $ 1725 "PSE_R≔pose_add(PSE_T, p[0,0,0.1,0,0,0])"
          global PSE_R= pose_add (PSE_T, p[0,0,0.1,0,0,0])
        end
      end
    end
    $ 1732 "Additional check"
    $ 1733 "If  not is_reachable(FRM_Reference,[PSE_A,PSE_A_H,PSE_T,PSE_T_H,PSE_R,PSE_R_H])"
    if (  not  is_reachable(FRM_Reference,[PSE_A,PSE_A_H,PSE_T,PSE_T_H,PSE_R,PSE_R_H])):
      $ 1734 "Error"
      $ 1735 "set_error(ERROR_POSE_NOT_REACHABLE)"
      set_error(ERROR_POSE_NOT_REACHABLE)
      $ 1736 "Action≔0"
      global Action=0
    end
    $ 1737 "'=========='"
    # '=========='
    $ 1738 "Switch Action"
    switch_1 = Action
    $ 1739 "Case 1"
    if (1 == switch_1):
      $ 1740 "Pick"
      $ 1741 "Action_Info≔'pick object'"
      global Action_Info="pick object"
      $ 1742 "do_transition(pose_trans(FRM_Reference, PSE_T), keep_rxry=OBJ_Picked)"
      do_transition( pose_trans (FRM_Reference, PSE_T), keep_rxry=OBJ_Picked)
      $ 1743 "EOAT"
      $ 1744 "If  not OBJ_Picked"
      if (  not  OBJ_Picked):
        $ 1745 "rq_move_and_wait_mm(GRP_Open_Pos)"
         rq_move_and_wait_mm (GRP_Open_Pos)
      end
      $ 1746 "If PSE_A_H≠PSE_Z"
      if (PSE_A_H != PSE_Z):
        $ 1747 "If JNT_Q≠JNT_Z"
        if (JNT_Q != JNT_Z):
          $ 1748 "movej(get_inverse_kin(pose_trans(FRM_Reference, PSE_A_H), qnear=JNT_Q), r=0.050)"
          movej(get_inverse_kin( pose_trans (FRM_Reference, PSE_A_H), qnear=JNT_Q), r=0.050)
        else:
          $ 1749 "Else" "noBreak"
          $ 1750 "movej(pose_trans(FRM_Reference, PSE_A_H), r=0.050)"
          movej( pose_trans (FRM_Reference, PSE_A_H), r=0.050)
        end
      end
      $ 1751 "If PSE_A≠PSE_Z"
      if (PSE_A != PSE_Z):
        $ 1752 "If JNT_Q≠JNT_Z"
        if (JNT_Q != JNT_Z):
          $ 1753 "movej(get_inverse_kin(pose_trans(FRM_Reference, PSE_A), qnear=JNT_Q), r=0.020)"
          movej(get_inverse_kin( pose_trans (FRM_Reference, PSE_A), qnear=JNT_Q), r=0.020)
        else:
          $ 1754 "Else" "noBreak"
          $ 1755 "movej(pose_trans(FRM_Reference, PSE_A), r=0.020)"
          movej( pose_trans (FRM_Reference, PSE_A), r=0.020)
        end
      end
      $ 1756 "MoveL"
      $ 1757 "If PSE_T_H≠PSE_Z"
      if (PSE_T_H != PSE_Z):
        $ 1758 "PSE_T_H" "breakAfter"
        movel(pose_trans(FRM_Reference, PSE_T_H), a=0.5, v=0.4, r=0.01)
      end
      $ 1759 "PSE_T" "breakAfter"
      movel(pose_trans(FRM_Reference, PSE_T), a=0.08, v=0.12)
      $ 1760 "EOAT"
      $ 1761 "rq_set_force_norm(50)"
       rq_set_force_norm (50)
      $ 1762 "rq_close_and_wait()"
       rq_close_and_wait ()
      $ 1763 "OBJ_Picked≔rq_is_object_detected()"
      global OBJ_Picked= rq_is_object_detected ()
      $ 1764 "If  not OBJ_Picked"
      if (  not  OBJ_Picked):
        $ 1765 "set_error(ERROR_NO_OBJECT_TO_PICK)"
        set_error(ERROR_NO_OBJECT_TO_PICK)
      end
      $ 1766 "EXTT"
      $ 1767 "Switch JIG"
      switch_2 = JIG
      $ 1768 "Case 1"
      if (1 == switch_2):
        $ 1769 "3FG"
        $ 1770 "If OBJ_Picked"
        if (OBJ_Picked):
          $ 1771 "Set GRP_3F_Open=On"
          set_standard_digital_out(5, True)
        end
      end
      $ 1772 "If PSE_R_H≠PSE_Z"
      if (PSE_R_H != PSE_Z):
        $ 1773 "PSE_R" "breakAfter"
        movel(pose_trans(FRM_Reference, PSE_R), a=0.5, v=0.4, r=0.01)
        $ 1774 "PSE_R_H" "breakAfter"
        movel(pose_trans(FRM_Reference, PSE_R_H), a=0.5, v=0.4)
      else:
        $ 1775 "Else" "noBreak"
        $ 1776 "PSE_R" "breakAfter"
        movel(pose_trans(FRM_Reference, PSE_R), a=0.5, v=0.4)
      end
    elif (2 == switch_1):
      $ 1777 "Case 2"
      $ 1778 "Place"
      $ 1779 "Action_Info≔'place object'"
      global Action_Info="place object"
      $ 1780 "do_transition(pose_trans(FRM_Reference, PSE_T), keep_rxry=OBJ_Picked)"
      do_transition( pose_trans (FRM_Reference, PSE_T), keep_rxry=OBJ_Picked)
      $ 1781 "EXTT"
      $ 1782 "Switch JIG"
      switch_2 = JIG
      $ 1783 "Case 1"
      if (1 == switch_2):
        $ 1784 "3FG"
        $ 1785 "If OBJ_Picked"
        if (OBJ_Picked):
          $ 1786 "Set GRP_3F_Open=On"
          set_standard_digital_out(5, True)
        end
      end
      $ 1787 "If PSE_A_H≠PSE_Z"
      if (PSE_A_H != PSE_Z):
        $ 1788 "If JNT_Q≠JNT_Z"
        if (JNT_Q != JNT_Z):
          $ 1789 "movej(get_inverse_kin(pose_trans(FRM_Reference, PSE_A_H), qnear=JNT_Q), r=0.050)"
          movej(get_inverse_kin( pose_trans (FRM_Reference, PSE_A_H), qnear=JNT_Q), r=0.050)
        else:
          $ 1790 "Else" "noBreak"
          $ 1791 "movej(pose_trans(FRM_Reference, PSE_A_H), r=0.050)"
          movej( pose_trans (FRM_Reference, PSE_A_H), r=0.050)
        end
      end
      $ 1792 "If PSE_A≠PSE_Z"
      if (PSE_A != PSE_Z):
        $ 1793 "If JNT_Q≠JNT_Z"
        if (JNT_Q != JNT_Z):
          $ 1794 "movej(get_inverse_kin(pose_trans(FRM_Reference, PSE_A), qnear=JNT_Q), r=0.020)"
          movej(get_inverse_kin( pose_trans (FRM_Reference, PSE_A), qnear=JNT_Q), r=0.020)
        else:
          $ 1795 "Else" "noBreak"
          $ 1796 "movej(pose_trans(FRM_Reference, PSE_A), r=0.020)"
          movej( pose_trans (FRM_Reference, PSE_A), r=0.020)
        end
      end
      $ 1797 "MoveL"
      $ 1798 "If PSE_T_H≠PSE_Z"
      if (PSE_T_H != PSE_Z):
        $ 1799 "PSE_T_H" "breakAfter"
        movel(pose_trans(FRM_Reference, PSE_T_H), a=0.5, v=0.4, r=0.01)
      end
      $ 1800 "PSE_T" "breakAfter"
      global move_thread_flag_1800=0
      thread move_thread_1800():
        enter_critical
        move_thread_flag_1800 = 1
        movel(pose_trans(FRM_Reference, PSE_T), a=0.05, v=0.09)
        move_thread_flag_1800 = 2
        exit_critical
      end
      move_thread_flag_1800 = 0
      move_thread_han_1800 = run move_thread_1800()
      while (True):
        local targetTcpDirection=get_target_tcp_speed()
        local stepsToRetract=tool_contact(direction=targetTcpDirection)
        if (stepsToRetract > 0):
          kill move_thread_han_1800
          stopl(0.5)
          $ 1801 "Until (tool_contact_detection)"
          break
        end
        sleep(1.0E-10)
        if (move_thread_flag_1800 > 1):
          join move_thread_han_1800
          break
        end
        sync()
      end
      $ 1802 "Force"
      sleep(0.02)
      zero_ftsensor()
      force_mode(FRM_Reference, [1, 1, 1, 0, 0, 0], [0.0, 0.0, 0.0, 0.0, 0.0, 0.0], 2, [0.1, 0.1, 0.01, 0.3490658503988659, 0.3490658503988659, 0.3490658503988659])
      $ 1803 "PSE_T" "noBreak"
      movel(pose_trans(FRM_Reference, PSE_T), a=0.04, v=0.07)
      end_force_mode()
      stopl(5.0)
      $ 1804 "EXTT"
      $ 1805 "Switch JIG"
      switch_2 = JIG
      $ 1806 "Case 1"
      if (1 == switch_2):
        $ 1807 "3FG"
        $ 1808 "If OBJ_Picked"
        if (OBJ_Picked):
          $ 1809 "Set GRP_3F_Open=Off"
          set_standard_digital_out(5, False)
          $ 1810 "Wait: 0.2"
          sleep(0.2)
        end
      end
      $ 1811 "EOAT"
      $ 1812 "rq_move_and_wait_mm(GRP_Open_Pos)"
       rq_move_and_wait_mm (GRP_Open_Pos)
      $ 1813 "OBJ_Picked≔rq_is_object_detected()"
      global OBJ_Picked= rq_is_object_detected ()
      $ 1814 "If PSE_R_H≠PSE_Z"
      if (PSE_R_H != PSE_Z):
        $ 1815 "PSE_R" "breakAfter"
        movel(pose_trans(FRM_Reference, PSE_R), a=0.5, v=0.4, r=0.01)
        $ 1816 "PSE_R_H" "breakAfter"
        movel(pose_trans(FRM_Reference, PSE_R_H), a=0.5, v=0.4)
      else:
        $ 1817 "Else" "noBreak"
        $ 1818 "PSE_R" "breakAfter"
        movel(pose_trans(FRM_Reference, PSE_R), a=0.5, v=0.4)
      end
    elif (3 == switch_1):
      $ 1819 "Case 3"
      $ 1820 "Push"
      $ 1821 "Action_Info≔'push'"
      global Action_Info="push"
    elif (4 == switch_1):
      $ 1822 "Case 4"
      $ 1823 "Pull"
      $ 1824 "Action_Info≔'pull'"
      global Action_Info="pull"
    elif (6 == switch_1):
      $ 1827 "Case 6"
      $ 1828 "Drop the cap"
      $ 1829 "If JNT_A≠[0,0,0,0,0,0]"
      if (JNT_A != [0,0,0,0,0,0]):
        $ 1830 "MoveJ"
        $ 1831 "JNT_A" "breakAfter"
        movej(JNT_A, a=1.3962634015954636, v=1.7453292519943295, r=0.02)
      else:
        $ 1832 "Else" "noBreak"
        $ 1833 "MoveJ"
        $ 1834 "PSE_A" "breakAfter"
        movej(pose_trans(FRM_Reference, PSE_A), a=1.3962634015954636, v=1.7453292519943295, r=0.02)
      end
      $ 1835 "MoveL"
      $ 1836 "PSE_T" "breakAfter"
      movel(pose_trans(FRM_Reference, PSE_T), a=0.05, v=0.09)
      $ 1837 "'ADD OPEN GRIPPER'"
      # 'ADD OPEN GRIPPER'
      # begin: URCap Program Node
      #   Source: Robotiq_Grippers, 3.17.0.105337, Robotiq Inc.
      #   Type: Gripper
      $ 1838 "Gripper Move10mm (1)"
      if not(gripper_connected[0]):
        popup("Gripper 1 must be connected to run this program.", "No connection", False, True, True)
      end
      if not(rq_is_gripper_activated("1")):
        popup("Gripper 1 is not activated. Go to Installation tab > Gripper to activate it and run the program again.", "Not activated", False, True, True)
      end
      rq_set_pos_spd_for(201, 0, 28, "1")
      rq_wait_pos_spe_for_request(201, 0, 28, "1")
      rq_go_to("1")
      rq_wait("1")
      # end: URCap Program Node
      $ 1839 "PSE_T_H" "breakAfter"
      movel(pose_trans(FRM_Reference, PSE_T_H), a=0.05, v=0.09)
      # begin: URCap Program Node
      #   Source: Robotiq_Grippers, 3.17.0.105337, Robotiq Inc.
      #   Type: Gripper
      $ 1840 "Gripper Move40mm (1)"
      if not(gripper_connected[0]):
        popup("Gripper 1 must be connected to run this program.", "No connection", False, True, True)
      end
      if not(rq_is_gripper_activated("1")):
        popup("Gripper 1 is not activated. Go to Installation tab > Gripper to activate it and run the program again.", "Not activated", False, True, True)
      end
      rq_set_pos_spd_for(63, 0, 28, "1")
      rq_wait_pos_spe_for_request(63, 0, 28, "1")
      rq_go_to("1")
      rq_wait("1")
      # end: URCap Program Node
      $ 1841 "PSE_R" "breakAfter"
      movel(pose_trans(FRM_Reference, PSE_R), a=0.5, v=0.4)
    elif (7 == switch_1):
      $ 1842 "Case 7"
      $ 1843 "Load"
      $ 1844 "Action_Info≔'load object'"
      global Action_Info="load object"
      $ 1845 "do_transition(pose_trans(FRM_Reference, PSE_T), keep_rxry=OBJ_Picked)"
      do_transition( pose_trans (FRM_Reference, PSE_T), keep_rxry=OBJ_Picked)
      $ 1846 "If PSE_A_H≠PSE_Z"
      if (PSE_A_H != PSE_Z):
        $ 1847 "If JNT_Q≠JNT_Z"
        if (JNT_Q != JNT_Z):
          $ 1848 "movej(get_inverse_kin(pose_trans(FRM_Reference, PSE_A_H), qnear=JNT_Q), r=0.050)"
          movej(get_inverse_kin( pose_trans (FRM_Reference, PSE_A_H), qnear=JNT_Q), r=0.050)
        else:
          $ 1849 "Else" "noBreak"
          $ 1850 "movej(pose_trans(FRM_Reference, PSE_A_H), r=0.050)"
          movej( pose_trans (FRM_Reference, PSE_A_H), r=0.050)
        end
      end
      $ 1851 "If PSE_A≠PSE_Z"
      if (PSE_A != PSE_Z):
        $ 1852 "If JNT_Q≠JNT_Z"
        if (JNT_Q != JNT_Z):
          $ 1853 "movej(get_inverse_kin(pose_trans(FRM_Reference, PSE_A), qnear=JNT_Q), r=0.020)"
          movej(get_inverse_kin( pose_trans (FRM_Reference, PSE_A), qnear=JNT_Q), r=0.020)
        else:
          $ 1854 "Else" "noBreak"
          $ 1855 "movej(pose_trans(FRM_Reference, PSE_A), r=0.020)"
          movej( pose_trans (FRM_Reference, PSE_A), r=0.020)
        end
      end
      $ 1856 "MoveL"
      $ 1857 "If PSE_T_H≠PSE_Z"
      if (PSE_T_H != PSE_Z):
        $ 1858 "PSE_T_H" "breakAfter"
        movel(pose_trans(FRM_Reference, PSE_T_H), a=0.5, v=0.4, r=0.01)
      end
      $ 1859 "PSE_T" "breakAfter"
      global move_thread_flag_1859=0
      thread move_thread_1859():
        enter_critical
        move_thread_flag_1859 = 1
        movel(pose_trans(FRM_Reference, PSE_T), a=0.05, v=0.09)
        move_thread_flag_1859 = 2
        exit_critical
      end
      move_thread_flag_1859 = 0
      move_thread_han_1859 = run move_thread_1859()
      while (True):
        local targetTcpDirection=get_target_tcp_speed()
        local stepsToRetract=tool_contact(direction=targetTcpDirection)
        if (stepsToRetract > 0):
          kill move_thread_han_1859
          stopl(0.5)
          $ 1860 "Until (tool_contact_detection)"
          break
        end
        sleep(1.0E-10)
        if (move_thread_flag_1859 > 1):
          join move_thread_han_1859
          break
        end
        sync()
      end
      $ 1861 "Force"
      sleep(0.02)
      zero_ftsensor()
      force_mode(FRM_Reference, [0, 1, 1, 0, 0, 1], [0.0, 0.0, 0.0, 0.0, 0.0, 0.0], 2, [0.1, 0.05, 0.02, 0.3490658503988659, 0.3490658503988659, 3.141592653589793])
      $ 1862 "PSE_T" "noBreak"
      movel(pose_trans(FRM_Reference, PSE_T), a=0.04, v=0.07)
      end_force_mode()
      stopl(5.0)
      $ 1863 "EOAT"
      $ 1864 "rq_move_and_wait_mm(GRP_Open_Pos)"
       rq_move_and_wait_mm (GRP_Open_Pos)
      $ 1865 "OBJ_Picked≔rq_is_object_detected()"
      global OBJ_Picked= rq_is_object_detected ()
      $ 1866 "If PSE_R_H≠PSE_Z"
      if (PSE_R_H != PSE_Z):
        $ 1867 "PSE_R" "breakAfter"
        movel(pose_trans(FRM_Reference, PSE_R), a=0.5, v=0.4, r=0.01)
        $ 1868 "PSE_R_H" "breakAfter"
        movel(pose_trans(FRM_Reference, PSE_R_H), a=0.5, v=0.4)
      else:
        $ 1869 "Else" "noBreak"
        $ 1870 "PSE_R" "breakAfter"
        movel(pose_trans(FRM_Reference, PSE_R), a=0.5, v=0.4)
      end
    elif (8 == switch_1):
      $ 1871 "Case 8"
      $ 1872 "Unload"
      $ 1873 "Action_Info≔'pick object'"
      global Action_Info="pick object"
      $ 1874 "do_transition(pose_trans(FRM_Reference, PSE_T), keep_rxry=OBJ_Picked)"
      do_transition( pose_trans (FRM_Reference, PSE_T), keep_rxry=OBJ_Picked)
      $ 1875 "EOAT"
      $ 1876 "If  not OBJ_Picked"
      if (  not  OBJ_Picked):
        $ 1877 "rq_move_and_wait_mm(GRP_Open_Pos)"
         rq_move_and_wait_mm (GRP_Open_Pos)
      end
      $ 1878 "If PSE_A_H≠PSE_Z"
      if (PSE_A_H != PSE_Z):
        $ 1879 "If JNT_Q≠JNT_Z"
        if (JNT_Q != JNT_Z):
          $ 1880 "movej(get_inverse_kin(pose_trans(FRM_Reference, PSE_A_H), qnear=JNT_Q), r=0.050)"
          movej(get_inverse_kin( pose_trans (FRM_Reference, PSE_A_H), qnear=JNT_Q), r=0.050)
        else:
          $ 1881 "Else" "noBreak"
          $ 1882 "movej(pose_trans(FRM_Reference, PSE_A_H), r=0.050)"
          movej( pose_trans (FRM_Reference, PSE_A_H), r=0.050)
        end
      end
      $ 1883 "If PSE_A≠PSE_Z"
      if (PSE_A != PSE_Z):
        $ 1884 "If JNT_Q≠JNT_Z"
        if (JNT_Q != JNT_Z):
          $ 1885 "movej(get_inverse_kin(pose_trans(FRM_Reference, PSE_A), qnear=JNT_Q), r=0.020)"
          movej(get_inverse_kin( pose_trans (FRM_Reference, PSE_A), qnear=JNT_Q), r=0.020)
        else:
          $ 1886 "Else" "noBreak"
          $ 1887 "movej(pose_trans(FRM_Reference, PSE_A), r=0.020)"
          movej( pose_trans (FRM_Reference, PSE_A), r=0.020)
        end
      end
      $ 1888 "MoveL"
      $ 1889 "If PSE_T_H≠PSE_Z"
      if (PSE_T_H != PSE_Z):
        $ 1890 "PSE_T_H" "breakAfter"
        movel(pose_trans(FRM_Reference, PSE_T_H), a=0.5, v=0.4, r=0.01)
      end
      $ 1891 "PSE_T" "breakAfter"
      movel(pose_trans(FRM_Reference, PSE_T), a=0.08, v=0.12)
      $ 1892 "Force"
      sleep(0.02)
      zero_ftsensor()
      force_mode(FRM_Reference, [1, 1, 0, 0, 0, 0], [0.0, 0.0, 0.0, 0.0, 0.0, 0.0], 2, [0.05, 0.05, 0.1, 0.3490658503988659, 0.3490658503988659, 0.3490658503988659])
      $ 1893 "EOAT" "noBreak"
      $ 1894 "rq_set_force_norm(50)" "noBreak"
       rq_set_force_norm (50)
      $ 1895 "rq_close_and_wait()" "noBreak"
       rq_close_and_wait ()
      $ 1896 "OBJ_Picked≔rq_is_object_detected()" "noBreak"
      global OBJ_Picked= rq_is_object_detected ()
      $ 1897 "If  not OBJ_Picked" "noBreak"
      if (  not  OBJ_Picked):
        $ 1898 "set_error(ERROR_NO_OBJECT_TO_PICK)" "noBreak"
        set_error(ERROR_NO_OBJECT_TO_PICK)
      end
      $ 1899 "If PSE_R_H≠PSE_Z" "noBreak"
      if (PSE_R_H != PSE_Z):
        $ 1900 "PSE_R" "noBreak"
        movel(pose_trans(FRM_Reference, PSE_R), a=0.5, v=0.4, r=0.01)
        $ 1901 "PSE_R_H" "noBreak"
        movel(pose_trans(FRM_Reference, PSE_R_H), a=0.5, v=0.4)
      else:
        $ 1902 "Else" "noBreak"
        $ 1903 "PSE_R" "noBreak"
        movel(pose_trans(FRM_Reference, PSE_R), a=0.5, v=0.4)
      end
      end_force_mode()
      stopl(5.0)
    elif (11 == switch_1):
      $ 1904 "Case 11"
    elif (12 == switch_1):
      $ 1941 "Case 12"
      $ 1942 "Decap"
      $ 1943 "Action_Info≔'decapping'"
      global Action_Info="decapping"
      $ 1944 "Set GRP_3F_Enable=On"
      set_standard_digital_out(4, True)
      $ 1945 "Set GRP_3F_Decap=On"
      set_standard_digital_out(3, True)
      $ 1946 "Force"
      sleep(0.02)
      zero_ftsensor()
      force_mode(tool_pose(), [0, 0, 1, 0, 0, 0], [0.0, 0.0, 5.0, 0.0, 0.0, 0.0], 2, [0.1, 0.1, 0.15, 0.3490658503988659, 0.3490658503988659, 0.3490658503988659])
      $ 1947 "check_decapping(offset=0.015, timeout=5, abort=CMD_Hold)" "noBreak"
      check_decapping(offset=0.015, timeout=5, abort=CMD_Hold)
      end_force_mode()
      stopl(5.0)
      $ 1948 "Set GRP_3F_Decap=Off"
      set_standard_digital_out(3, False)
      $ 1949 "Set GRP_3F_Enable=Off"
      set_standard_digital_out(4, False)
      $ 1950 "MoveL"
      $ 1951 "PSE_R" "breakAfter"
      movel(pose_trans(FRM_Reference, PSE_R), a=0.8, v=0.15)
    elif (13 == switch_1):
      $ 1952 "Case 13"
      $ 1953 "TMR_Barcode: Reset"
      TMR_Barcode = 0
      $ 1954 "Read"
      $ 1955 "TMR_Barcode: Start"
      TMR_Barcode_is_counting = True
      $ 1956 "If TMR_Barcode<PRM_TO_Read_BC"
      global thread_flag_1956=0
      thread Thread_if_1956():
        $ 1957 "KeyenceTrigger"
        $ 1958 "Set OClearResult=HI:Pulse 0.2"
        thread SinglePulse98():
          write_output_boolean_register(2, True)
          sleep(0.2)
          write_output_boolean_register(2, False)
        end
        singlePulse98 = run SinglePulse98()
        $ 1959 "Wait: 0.5"
        sleep(0.5)
        $ 1960 "Set OTriggerBarcode=Off"
        write_output_boolean_register(1, False)
        $ 1961 "Wait: 0.5"
        sleep(0.5)
        $ 1962 "Set OTriggerBarcode=On"
        write_output_boolean_register(1, True)
        $ 1963 "Wait: 0.5"
        sleep(0.5)
        $ 1964 "Preorient"
        $ 1965 "TMR_Barcode: Reset"
        TMR_Barcode = 0
        $ 1966 "If ICmdExctd"
        if (read_input_boolean_register(12)):
          $ 1967 "Set GRP_3F_Decap=On"
          set_standard_digital_out(3, True)
          $ 1968 "Set GRP_3F_Enable=On"
          set_standard_digital_out(4, True)
          $ 1969 "Loop ICmdExctd"
          while (read_input_boolean_register(12)):
            $ 1970 "KeyenceTrigger"
            $ 1971 "Set OClearResult=HI:Pulse 0.1"
            thread SinglePulse99():
              write_output_boolean_register(2, True)
              sleep(0.1)
              write_output_boolean_register(2, False)
            end
            singlePulse99 = run SinglePulse99()
            $ 1972 "Wait: 0.3"
            sleep(0.3)
            $ 1973 "Set OTriggerBarcode=Off"
            write_output_boolean_register(1, False)
            $ 1974 "Wait: 0.3"
            sleep(0.3)
            $ 1975 "Set OTriggerBarcode=On"
            write_output_boolean_register(1, True)
            $ 1976 "Wait: 0.1"
            sleep(0.1)
          end
        end
        $ 1977 "If  not ICmdExctd"
        if (  not  read_input_boolean_register(12)):
          $ 1978 "Set GRP_3F_Decap=On"
          set_standard_digital_out(3, True)
          $ 1979 "Set GRP_3F_Enable=On"
          set_standard_digital_out(4, True)
          $ 1980 "Wait ICmdExctd=HI"
          while (read_input_boolean_register(12) == False):
            sync()
          end
        end
        $ 1981 "Set GRP_3F_Decap=Off"
        set_standard_digital_out(3, False)
        $ 1982 "Set GRP_3F_Enable=Off"
        set_standard_digital_out(4, False)
        $ 1983 "OBJ_Brc_OK≔ True "
        global OBJ_Brc_OK=  True
        thread_flag_1956 = 1
      end
      if (TMR_Barcode<PRM_TO_Read_BC):
        global thread_handler_1956=run Thread_if_1956()
        while (thread_flag_1956 == 0):
          if not(TMR_Barcode<PRM_TO_Read_BC):
            kill thread_handler_1956
            thread_flag_1956 = 2
          else:
            sync()
          end
        end
      else:
        thread_flag_1956 = 2
      end
      if (thread_flag_1956 == 2):
        $ 1984 "Else" "noBreak"
        $ 1985 "exeption"
        $ 1986 "error"
        $ 1988 "OBJ_Brc_OK≔ False "
        global OBJ_Brc_OK=  False
      end
      $ 1989 "Set GRP_3F_Decap=Off"
      set_standard_digital_out(3, False)
      $ 1990 "Set GRP_3F_Enable=Off"
      set_standard_digital_out(4, False)
      $ 1991 "Set OTriggerBarcode=Off"
      write_output_boolean_register(1, False)
    elif (15 == switch_1):
      $ 1992 "Case 15"
      $ 1993 "Detect"
      $ 1994 "Action_Info≔'detect'"
      global Action_Info="detect"
    elif (30 == switch_1):
      $ 1995 "Case 30"
      $ 1996 "Shake"
      $ 1997 "Action_Info≔'shake'"
      global Action_Info="shake"
      $ 1998 "do_transition(pose_trans(FRM_Reference, PSE_T), keep_rxry=OBJ_Picked)"
      do_transition( pose_trans (FRM_Reference, PSE_T), keep_rxry=OBJ_Picked)
      $ 1999 "If PSE_A_H≠PSE_Z"
      if (PSE_A_H != PSE_Z):
        $ 2000 "If JNT_Q≠JNT_Z"
        if (JNT_Q != JNT_Z):
          $ 2001 "movej(get_inverse_kin(pose_trans(FRM_Reference, PSE_A_H), qnear=JNT_Q), r=0.050)"
          movej(get_inverse_kin( pose_trans (FRM_Reference, PSE_A_H), qnear=JNT_Q), r=0.050)
        else:
          $ 2002 "Else" "noBreak"
          $ 2003 "movej(pose_trans(FRM_Reference, PSE_A_H), r=0.050)"
          movej( pose_trans (FRM_Reference, PSE_A_H), r=0.050)
        end
      end
      $ 2004 "If PSE_A≠PSE_Z"
      if (PSE_A != PSE_Z):
        $ 2005 "If JNT_Q≠JNT_Z"
        if (JNT_Q != JNT_Z):
          $ 2006 "movej(get_inverse_kin(pose_trans(FRM_Reference, PSE_A), qnear=JNT_Q), r=0.020)"
          movej(get_inverse_kin( pose_trans (FRM_Reference, PSE_A), qnear=JNT_Q), r=0.020)
        else:
          $ 2007 "Else" "noBreak"
          $ 2008 "movej(pose_trans(FRM_Reference, PSE_A), r=0.020)"
          movej( pose_trans (FRM_Reference, PSE_A), r=0.020)
        end
      end
      $ 2009 "MoveL"
      $ 2010 "If PSE_T_H≠PSE_Z"
      if (PSE_T_H != PSE_Z):
        $ 2011 "PSE_T_H" "breakAfter"
        movel(pose_trans(FRM_Reference, PSE_T_H), a=0.5, v=0.4, r=0.01)
      end
      $ 2012 "PSE_T" "breakAfter"
      movel(pose_trans(FRM_Reference, PSE_T), a=0.08, v=0.12)
      $ 2013 "EXTT"
      $ 2014 "Comment"
      # Comment
      $ 2015 "MoveJ"
      $ 2016 "Waypoint_54" "breakAfter"
      movej(get_inverse_kin(Waypoint_54_p, qnear=Waypoint_54_q), a=1.3962634015954636, v=1.0471975511965976)
      $ 2017 "MoveJ"
      $ 2018 "Waypoint_77" "breakAfter"
      movej(get_inverse_kin(Waypoint_77_p, qnear=Waypoint_77_q), a=1.3962634015954636, v=1.0471975511965976)
      $ 2019 "MoveJ"
      $ 2020 "Waypoint_83" "breakAfter"
      movej(get_inverse_kin(Waypoint_83_p, qnear=Waypoint_83_q), a=1.3962634015954636, v=1.0471975511965976)
      $ 2021 "MoveJ"
      $ 2022 "Waypoint_84" "breakAfter"
      movej(get_inverse_kin(Waypoint_84_p, qnear=Waypoint_84_q), a=1.3962634015954636, v=1.0471975511965976)
      $ 2023 "If PSE_R_H≠PSE_Z"
      if (PSE_R_H != PSE_Z):
        $ 2024 "PSE_R" "breakAfter"
        movel(pose_trans(FRM_Reference, PSE_R), a=0.5, v=0.4, r=0.01)
        $ 2025 "PSE_R_H" "breakAfter"
        movel(pose_trans(FRM_Reference, PSE_R_H), a=0.5, v=0.4)
      else:
        $ 2026 "Else" "noBreak"
        $ 2027 "PSE_R" "breakAfter"
        movel(pose_trans(FRM_Reference, PSE_R), a=0.5, v=0.4)
      end
    elif (31 == switch_1):
      $ 2028 "Case 31"
      $ 2029 "Action_Info≔'Pick_Vial'"
      global Action_Info="Pick_Vial"
      $ 2030 "Pick_Vial"
      # begin: URCap Program Node
      #   Source: Robotiq_Grippers, 3.17.0.105337, Robotiq Inc.
      #   Type: Gripper
      $ 2031 "Gripper Open (1)"
      if not(gripper_connected[0]):
        popup("Gripper 1 must be connected to run this program.", "No connection", False, True, True)
      end
      if not(rq_is_gripper_activated("1")):
        popup("Gripper 1 is not activated. Go to Installation tab > Gripper to activate it and run the program again.", "Not activated", False, True, True)
      end
      rq_set_pos_spd_for(0, 82, 71, "1")
      rq_wait_pos_spe_for_request(0, 82, 71, "1")
      rq_go_to("1")
      rq_wait("1")
      # end: URCap Program Node
      $ 2032 "MoveJ"
      $ 2033 "Vial_above_1" "breakAfter"
      movej(get_inverse_kin(Vial_above_1_p, qnear=Vial_above_1_q), a=0.5235987755982988, v=0.4363323129985824, r=0.05)
      $ 2034 "MoveL"
      $ 2035 "Vial_pick_poi_1" "breakAfter"
      movel(Vial_pick_poi_1_p, a=0.5, v=0.1)
      # begin: URCap Program Node
      #   Source: Robotiq_Grippers, 3.17.0.105337, Robotiq Inc.
      #   Type: Gripper
      $ 2036 "Gripper Close (1)"
      if not(gripper_connected[0]):
        popup("Gripper 1 must be connected to run this program.", "No connection", False, True, True)
      end
      if not(rq_is_gripper_activated("1")):
        popup("Gripper 1 is not activated. Go to Installation tab > Gripper to activate it and run the program again.", "Not activated", False, True, True)
      end
      rq_set_pos_spd_for(255, 71, 84, "1")
      rq_wait_pos_spe_for_request(255, 71, 84, "1")
      rq_go_to("1")
      rq_wait("1")
      # end: URCap Program Node
      $ 2037 "MoveL"
      $ 2038 "Waypoint_86" "breakAfter"
      movel(Waypoint_86_p, a=0.5, v=0.1, r=0.05)
      $ 2039 "Home (Safe)"
      movej([-1.2302089344500047, -1.2969853503591224, -1.875639182904262, -1.539621866126728, 1.5731943360401213, -2.80099559440227], a=1.3962634015954636, v=1.0471975511965976)
    elif (32 == switch_1):
      $ 2040 "Case 32"
      $ 2042 "decap_Vial"
      $ 2043 "Set GRP_3F_Open=On"
      set_standard_digital_out(5, True)
      $ 2044 "MoveJ"
      $ 2045 "Waypoint_87" "breakAfter"
      movej(get_inverse_kin(Waypoint_87_p, qnear=Waypoint_87_q), a=0.5235987755982988, v=0.4363323129985824)
      $ 2046 "MoveL"
      $ 2047 "Vial_3FG_plac_1" "breakAfter"
      movel(Vial_3FG_plac_1_p, a=0.5, v=0.1)
      $ 2048 "Set GRP_3F_Open=Off"
      set_standard_digital_out(5, False)
      $ 2049 "Wait: 0.5"
      sleep(0.5)
      $ 2050 "MoveL"
      $ 2051 "Waypoint_88" "breakAfter"
      movel(Waypoint_88_p, a=0.5, v=0.1, r=0.05)
      $ 2052 "MoveJ"
      $ 2053 "cap_dump_1" "breakAfter"
      movej(get_inverse_kin(cap_dump_1_p, qnear=cap_dump_1_q), a=0.5235987755982988, v=0.4363323129985824)
      # begin: URCap Program Node
      #   Source: Robotiq_Grippers, 3.17.0.105337, Robotiq Inc.
      #   Type: Gripper
      $ 2054 "Gripper Open (1)"
      if not(gripper_connected[0]):
        popup("Gripper 1 must be connected to run this program.", "No connection", False, True, True)
      end
      if not(rq_is_gripper_activated("1")):
        popup("Gripper 1 is not activated. Go to Installation tab > Gripper to activate it and run the program again.", "Not activated", False, True, True)
      end
      rq_set_pos_spd_for(0, 255, 255, "1")
      rq_wait_pos_spe_for_request(0, 255, 255, "1")
      rq_go_to("1")
      rq_wait("1")
      # end: URCap Program Node
      $ 2055 "MoveJ"
      $ 2056 "Waypoint_89" "breakAfter"
      movej(get_inverse_kin(Waypoint_89_p, qnear=Waypoint_89_q), a=0.5235987755982988, v=0.4363323129985824, r=0.05)
      $ 2057 "MoveL"
      $ 2058 "Vial_3FG_plac_2" "breakAfter"
      movel(Vial_3FG_plac_2_p, a=0.5, v=0.1)
      # begin: URCap Program Node
      #   Source: Robotiq_Grippers, 3.17.0.105337, Robotiq Inc.
      #   Type: Gripper
      $ 2059 "Gripper Close (1)"
      if not(gripper_connected[0]):
        popup("Gripper 1 must be connected to run this program.", "No connection", False, True, True)
      end
      if not(rq_is_gripper_activated("1")):
        popup("Gripper 1 is not activated. Go to Installation tab > Gripper to activate it and run the program again.", "Not activated", False, True, True)
      end
      rq_set_pos_spd_for(255, 204, 255, "1")
